   // ---- GENERATED: setup
   IF #Startup OR NOT #Core.Named THEN
       #InstancePath := GetInstancePath(size := 0);
       "FRK_SetIdentity"(Core := #Core,
                         Status := #Status,
                         InstancePath := #InstancePath,
                         ModuleType := 1,
                         TypeId := 4,
                         Capabilities := DWORD#16#00000000,
                         ParentIndex := #ParentIndex,
                         TypeKey := 'Fraktal.Test.Satellite');
   END_IF;
   IF #Startup OR #ConfigRev = 0 THEN
       #ConfigRev := "FRK_ConfigRevision"(Previous := #ConfigRev);
   END_IF;
   #SupportedModesPublished[0] := TRUE;
   #SupportedModesPublished[1] := TRUE;
   #SupportedModesPublished[2] := TRUE;
   #SupportedModesPublished[3] := FALSE;
   #SupportedModesPublished[4] := FALSE;
   #SupportedModesPublished[5] := FALSE;
   #SupportedModesPublished[6] := FALSE;
   "FRK_UnitPrepare"(Core := #Core,
                     Unit := #Unit,
                     Policy := #ModePolicy,
                     Request := #HmiRequest,
                     Response := #HmiResponse,
                     Startup := #Startup,
                     InitialMode := 1);
   "FRK_AccessCyclic"(Access := #Access,
                      Startup := #Startup,
                      SourcePath := STRING_TO_WSTRING(#Status.Name),
                      History := #History,
                      Head := #HistoryHead,
                      Revision := #ConfigRev);
   "FRK_UnitMailbox"(Core := #Core,
                     Unit := #Unit,
                     Status := #Status,
                     Policy := #ModePolicy,
                     Access := #Access,
                     Request := #HmiRequest,
                     Response := #HmiResponse,
                     Supported := #SupportedModesPublished);
   // ---- GENERATED: begin
   "FRK_Begin"(Core := #Core,
               Status := #Status,
               Execute := #Unit.RunReq,
               Abort := (#Abort OR #Unit.AbortReq),
               Command := 1);
   IF #Core.EvCommandStart THEN
       #LatchedParCmd := #ParCmd;
       CASE #Core.Command OF
           1:
               "FRK_UnitRunStart"(Core := #Core,
                                  Status := #Status,
                                  Timeout := #ParCfg.Timeout,
                                  Label := 'Run');
           ELSE
               "FRK_Start"(Core := #Core,
                           Status := #Status,
                           Supported := FALSE,
                           Timeout := T#0ms,
                           Label := '');
       END_CASE;
   END_IF;
   IF #Core.EvCommandStart THEN
       // ---- AUTHORED: CommandStart
       #Device.Received := "FRK_PartReceived"(Core := #Core, Unit := #Unit, Status := #Status, Part := #Part, History := #History, Head := #HistoryHead);
       IF #Device.Received THEN
           "FRK_PartStarted"(Unit := #Unit,
                             Status := #Status,
                             Part := #Part,
                             History := #History,
                             Head := #HistoryHead);
       END_IF;
       // ---- GENERATED: reaction end
   END_IF;
   // ---- AUTHORED: cyclic management
   IF #Hal.Cell.Clamp.BackgroundFault THEN
       "FRK_Fault"(Core := #Core,
                   Status := #Status,
                   ReasonCode := 2901,
                   Description := WSTRING#'test.unit.condition');
   END_IF;
   // ---- GENERATED: end management
   "FRK_Release_SatelliteUnit"(Unit := #Unit,
                               Hal := #Hal);
   "FRK_UnitConsume"(Core := #Core,
                     Unit := #Unit,
                     Status := #Status,
                     Policy := #ModePolicy,
                     Access := #Access,
                     Response := #HmiResponse,
                     Supported := #SupportedModesPublished);
   "FRK_UnitMode"(Core := #Core,
                  Unit := #Unit);
   IF #Core.EvModeExit THEN
       // ---- AUTHORED: ModeExit
       #Device.ExitCalls := #Device.ExitCalls + 1;
       IF #Hal.Cell.Clamp.ExitHold THEN
           #Core.HookResult := 1;
       ELSE
           #Core.HookResult := 0;
       END_IF;
       // ---- GENERATED: reaction end
   END_IF;
   "FRK_UnitModeResolve"(Core := #Core,
                         Unit := #Unit,
                         Status := #Status,
                         Policy := #ModePolicy,
                         Timeout := #ParCfg.Timeout);
   IF #Core.EvModeChanged THEN
       // ---- AUTHORED: ModeChanged
       #Device.Changes := #Device.Changes + 1;
       // ---- GENERATED: reaction end
   END_IF;
   "FRK_UnitFollow"(Core := #Core,
                    Unit := #Unit,
                    Status := #Status,
                    Policy := #ModePolicy,
                    Access := #Access,
                    Supported := #SupportedModesPublished);
   IF #Unit.RequestPending AND (#Unit.Request.Kind = 11 OR #Unit.Request.Kind = 16) THEN
       #ManualMatched := FALSE;
       #RouteMatched := "FRK_Route_DeclarationCell"(Module := #Cell, Hal := #Hal.Cell, Request := #Unit.Request, Report := #HmiResponse.Report);
       #ManualMatched := #ManualMatched OR #RouteMatched;
       #RouteMatched := "FRK_Route_InnerUnit"(Module := #Inner, Hal := #Hal.Inner, Request := #Unit.Request, Report := #HmiResponse.Report);
       #ManualMatched := #ManualMatched OR #RouteMatched;
       IF NOT #ManualMatched THEN
           "FRK_ReleaseReason"(Report := #HmiResponse.Report,
                               Description := WSTRING#'std.error.unsupportedHmiRequest',
                               Reason := 2008,
                               Path := #Unit.Request.TargetPath,
                               Kind := 4);
       END_IF;
       #HmiResponse.Accepted := #Unit.Request.Kind = 16 OR #HmiResponse.Report.Released;
       IF #Unit.Request.Kind = 11 THEN
           IF #HmiResponse.Accepted THEN
               #HmiResponse.Diagnostic := WSTRING#'std.audit.manualCommandAccepted';
           ELSE
               #HmiResponse.Diagnostic := WSTRING#'std.audit.manualCommandRejected';
           END_IF;
       END_IF;
   END_IF;
   IF #Unit.EvReset THEN
       // ---- AUTHORED: OperatorReset
       #Device.Resets := #Device.Resets + 1;
       // ---- GENERATED: reset reaction end
   END_IF;
   IF #Core.ReleasePending OR #Unit.ReleaseChildren THEN
       "FRK_ReleaseCommand"(Core := #Cell.Core,
                            Execute := #Cell.Execute);
       "FRK_ReleaseCommand"(Core := #Inner.Core,
                            Execute := #Inner.Execute);
   END_IF;
   // ---- GENERATED: child call
   #Cell(ParentIndex := #Core.RegIndex,
         Startup := #Startup,
         Hal := #Hal.Cell);
   "FRK_ManualFinish"(Core := #Cell.Core,
                      Execute := #Cell.Execute,
                      ManualOwned := #Cell.ManualOwned);
   "FRK_UnitCascade"(ParentUnit := #Unit,
                     Core := #Inner.Core,
                     Unit := #Inner.Unit,
                     Status := #Inner.Status,
                     Policy := #Inner.ModePolicy,
                     Access := #Inner.Access,
                     Supported := #Inner.SupportedModesPublished,
                     History := #History,
                     Head := #HistoryHead);
   // ---- GENERATED: child call
   #Inner(ParentIndex := #Core.RegIndex,
          Startup := #Startup,
          Hal := #Hal.Inner);
   #Unit.CascadePending := FALSE;
   IF #Unit.RequestPending AND #Unit.Request.Kind = 23 THEN
       #HmiResponse.Accepted := FALSE;
       #HmiResponse.Report.Count := 0;
       #HmiResponse.Report.Released := TRUE;
       #HmiResponse.Diagnostic := WSTRING#'';
       "FRK_ConfigBegin"(Cursor := #ConfigCursor,
                         Page := #HmiResponse.ConfigPage,
                         PageIndex := #Unit.Request.IntValue,
                         Revision := #ConfigRev);
       IF #Unit.Request.DurationMs <> 0 THEN
           #HmiResponse.Diagnostic := WSTRING#'std.error.modelNotAvailable';
       ELSIF #Unit.Request.IntValue < 0 OR #Unit.Request.IntValue > 32767 THEN
           #HmiResponse.Diagnostic := WSTRING#'std.error.hmiRequestRejected';
       ELSE
           "FRK_ConfigUnit"(Scope := #Status.Name,
                            Policy := #ModePolicy,
                            ReadLevel := #Access.Policy.Required[0],
                            Readable := #Access.CurrentLevel >= #Access.Policy.Required[0],
                            Cursor := #ConfigCursor,
                            Page := #HmiResponse.ConfigPage);
           "FRK_Config_DeclarationCell"(Module := #Cell,
                                        ReadLevel := #Access.Policy.Required[0],
                                        Readable := #Access.CurrentLevel >= #Access.Policy.Required[0],
                                        Cursor := #ConfigCursor,
                                        Page := #HmiResponse.ConfigPage);
           "FRK_Config_InnerUnit"(Module := #Inner,
                                  ReadLevel := #Access.Policy.Required[0],
                                  Readable := #Access.CurrentLevel >= #Access.Policy.Required[0],
                                  Cursor := #ConfigCursor,
                                  Page := #HmiResponse.ConfigPage);
           "FRK_ConfigFinish"(Cursor := #ConfigCursor,
                              Page := #HmiResponse.ConfigPage);
           #HmiResponse.Accepted := TRUE;
       END_IF;
   END_IF;
   "FRK_RouteAbort"(Core := #Core,
                    Abort := (#Abort OR #Unit.AbortReq));
   IF #Core.EvAbort THEN
       "FRK_PartAborted"(Core := #Core,
                         Unit := #Unit,
                         Status := #Status,
                         Part := #Part,
                         History := #History,
                         Head := #HistoryHead);
   END_IF;
   IF #Core.Dispatch AND #Core.RegIndex > 0 AND NOT "FRK_Registry".Fault THEN
       // ---- AUTHORED: dispatch
       IF #Hal.Cell.Clamp.Finish THEN
           #Device.Processed := FALSE;
           IF #Unit.CarrierIndex = 0 THEN
               #Device.Processed := TRUE;
           ELSE
               #Device.Processed := "FRK_PartProcessed"(Core := #Core, Unit := #Unit, Status := #Status, Part := #Part, History := #History, Head := #HistoryHead, Verdict := #Hal.Cell.Clamp.Verdict, Reason := #Hal.Cell.Clamp.Diag.ReasonCode);
           END_IF;
           IF #Device.Processed THEN
               #Device.Cycles := #Device.Cycles + 1;
               IF #Unit.StopReq THEN
                   "FRK_Complete"(Core := #Core,
                                  Status := #Status);
               ELSE
                   #Device.Received := "FRK_PartReceived"(Core := #Core, Unit := #Unit, Status := #Status, Part := #Part, History := #History, Head := #HistoryHead);
                   IF #Device.Received THEN
                       "FRK_PartStarted"(Unit := #Unit,
                                         Status := #Status,
                                         Part := #Part,
                                         History := #History,
                                         Head := #HistoryHead);
                   END_IF;
               END_IF;
           END_IF;
       END_IF;
       // ---- GENERATED: end dispatch
   END_IF;
   "FRK_End"(Core := #Core,
             Status := #Status,
             Busy => #Busy,
             Done => #Done,
             Error => #Error,
             Aborted => #Aborted,
             Held => #Held,
             ErrorID => #ErrorID,
             Timing => #Timing);
   "FRK_AccessFinish"(Access := #Access,
                      Unit := #Unit,
                      Response := #HmiResponse,
                      SourcePath := STRING_TO_WSTRING(#Status.Name),
                      History := #History,
                      Head := #HistoryHead,
                      Revision := #ConfigRev);
   "FRK_UnitFinish"(Core := #Core,
                    Unit := #Unit,
                    Response := #HmiResponse,
                    Status := #Status,
                    Part := #Part,
                    History := #History,
                    Head := #HistoryHead);
   #ModeActivePublished := #Unit.Mode;
   #RunningPublished := #Core.Exec = 1;
   #StopPendingPublished := #Unit.StopReq AND #Core.Exec = 1;
   #GoodCount := #Unit.Good;
   #NokCount := #Unit.Nok;
   #ReworkCount := #Unit.Rework;
   #NokReason := #Unit.NokReason;
   // ---- AUTHORED: unconditional cyclic/derived data
   #OutImm.Cycles := #Device.Cycles;
   #OutImm.ExitCalls := #Device.ExitCalls;
   #OutImm.Changes := #Device.Changes;
   #OutImm.Resets := #Device.Resets;
   // ---- GENERATED: frame end
END_FUNCTION_BLOCK

FUNCTION_BLOCK "FB_InnerUnit"   // FB3, SCL
{ S7_Optimized_Access := 'TRUE' }
VERSION : 0.1
// Generated frame v0.6; change the declaration, then regenerate.
// stored: AutoNumber true, IsIECCheckEnabled false, IsRetainMemResEnabled false, MemoryReserve 100, SetENOAutomatically false, UDAEnableTagReadback false
   VAR_INPUT
      Execute { ExternalWritable := 'False'} : Bool;
      Abort { ExternalWritable := 'False'} : Bool;
      Command { ExternalWritable := 'False'} : DInt;
      ParCfg { ExternalWritable := 'False'} : "ST_DeclarationParCfg";
      ParCmd { ExternalWritable := 'False'} : "ST_DeclarationParCmd";
      ParentIndex { ExternalAccessible := 'False'; ExternalVisible := 'False'; ExternalWritable := 'False'} : DInt;
      Startup { ExternalAccessible := 'False'; ExternalVisible := 'False'; ExternalWritable := 'False'} : Bool;
   END_VAR
   VAR_OUTPUT
      Busy { ExternalWritable := 'False'} : Bool;
      Done { ExternalWritable := 'False'} : Bool;
      Error { ExternalWritable := 'False'} : Bool;
      Aborted { ExternalWritable := 'False'} : Bool;
      Held { ExternalWritable := 'False'} : Bool;
      ErrorID { ExternalWritable := 'False'} : DWord;
      Timing { ExternalWritable := 'False'} : "ST_ModuleTiming";
      OutCmd { ExternalWritable := 'False'} : "ST_DeclarationOutCmd";
      OutImm { ExternalWritable := 'False'} : "ST_UnitProbeImm";
   END_VAR
   VAR_IN_OUT
      Hal : "ST_InnerUnitHal";
   END_VAR
   VAR
      Status { ExternalWritable := 'False'; S7_SetPoint := 'True'} : "ST_ModuleStatus";
      Core { ExternalAccessible := 'False'; ExternalVisible := 'False'; ExternalWritable := 'False'; S7_SetPoint := 'True'} : "FRK_Core";
      LatchedParCmd { ExternalAccessible := 'False'; ExternalVisible := 'False'; ExternalWritable := 'False'; S7_SetPoint := 'True'} : "ST_DeclarationParCmd";
      Device { ExternalAccessible := 'False'; ExternalVisible := 'False'; ExternalWritable := 'False'; S7_SetPoint := 'True'} : "ST_UnitProbeDevice";
      Unit { ExternalAccessible := 'False'; ExternalVisible := 'False'; ExternalWritable := 'False'; S7_SetPoint := 'True'} : "FRK_Unit";
      HmiRequest { S7_SetPoint := 'True'} : "ST_HmiRequest";
      ModePolicy { ExternalAccessible := 'False'; ExternalVisible := 'False'; ExternalWritable := 'False'; S7_SetPoint := 'True'} : Array[0..6] of "ST_ModePolicy";
      Access { ExternalWritable := 'False'; S7_SetPoint := 'True'} : "FRK_Access";
      HmiResponse { ExternalWritable := 'False'; S7_SetPoint := 'True'} : "ST_HmiResponse";
      ConfigRev { ExternalWritable := 'False'} : UDInt;
      ConfigCursor { ExternalAccessible := 'False'; ExternalVisible := 'False'; ExternalWritable := 'False'; S7_SetPoint := 'True'} : "FRK_ConfigCursor";
      Part { ExternalWritable := 'False'; S7_SetPoint := 'True'} : "ST_PartContext";
      History { ExternalWritable := 'False'; S7_SetPoint := 'True'} : Array[1..16] of "ST_Diagnostic";
      HistoryHead { ExternalWritable := 'False'} : Int;
      ModeActivePublished { ExternalWritable := 'False'} : DInt;
      RunningPublished { ExternalWritable := 'False'} : Bool;
      StopPendingPublished { ExternalWritable := 'False'} : Bool;
      SupportedModesPublished { ExternalWritable := 'False'} : Array[0..6] of Bool;
      GoodCount { ExternalWritable := 'False'} : UDInt;
      NokCount { ExternalWritable := 'False'} : UDInt;
      ReworkCount { ExternalWritable := 'False'} : UDInt;
      NokReason { ExternalWritable := 'False'} : DInt;
      Cell { ExternalWritable := 'False'; S7_SetPoint := 'True'} : "FB_DeclarationCell";
   END_VAR
   VAR_TEMP
      InstancePath : WString[254];
      RouteMatched : Bool;
      ManualMatched : Bool;
   END_VAR
   VAR CONSTANT
      EXEC_READY : DInt := 0;
      MODULE_TIER : DInt := 1;
   END_VAR
BEGIN

   // ---- GENERATED: setup
   IF #Startup OR NOT #Core.Named THEN
       #InstancePath := GetInstancePath(size := 0);
       "FRK_SetIdentity"(Core := #Core,
                         Status := #Status,
                         InstancePath := #InstancePath,
                         ModuleType := 1,
                         TypeId := 5,
                         Capabilities := DWORD#16#00000000,
                         ParentIndex := #ParentIndex,
                         TypeKey := 'Fraktal.Test.Inner');
   END_IF;
   IF #Startup OR #ConfigRev = 0 THEN
       #ConfigRev := "FRK_ConfigRevision"(Previous := #ConfigRev);
   END_IF;
   #SupportedModesPublished[0] := TRUE;
   #SupportedModesPublished[1] := TRUE;
   #SupportedModesPublished[2] := TRUE;
   #SupportedModesPublished[3] := FALSE;
   #SupportedModesPublished[4] := FALSE;
   #SupportedModesPublished[5] := FALSE;
   #SupportedModesPublished[6] := FALSE;
   "FRK_UnitPrepare"(Core := #Core,
                     Unit := #Unit,
                     Policy := #ModePolicy,
                     Request := #HmiRequest,
                     Response := #HmiResponse,
                     Startup := #Startup,
                     InitialMode := 1);
   "FRK_AccessCyclic"(Access := #Access,
                      Startup := #Startup,
                      SourcePath := STRING_TO_WSTRING(#Status.Name),
                      History := #History,
                      Head := #HistoryHead,
                      Revision := #ConfigRev);
   "FRK_UnitMailbox"(Core := #Core,
                     Unit := #Unit,
                     Status := #Status,
                     Policy := #ModePolicy,
                     Access := #Access,
                     Request := #HmiRequest,
                     Response := #HmiResponse,
                     Supported := #SupportedModesPublished);
   // ---- GENERATED: begin
   "FRK_Begin"(Core := #Core,
               Status := #Status,
               Execute := #Unit.RunReq,
               Abort := (#Abort OR #Unit.AbortReq),
               Command := 1);
   IF #Core.EvCommandStart THEN
       #LatchedParCmd := #ParCmd;
       CASE #Core.Command OF
           1:
               "FRK_UnitRunStart"(Core := #Core,
                                  Status := #Status,
                                  Timeout := #ParCfg.Timeout,
                                  Label := 'Run');
           ELSE
               "FRK_Start"(Core := #Core,
                           Status := #Status,
                           Supported := FALSE,
                           Timeout := T#0ms,
                           Label := '');
       END_CASE;
   END_IF;
   IF #Core.EvCommandStart THEN
       // ---- AUTHORED: CommandStart
       #Device.Received := "FRK_PartReceived"(Core := #Core, Unit := #Unit, Status := #Status, Part := #Part, History := #History, Head := #HistoryHead);
       IF #Device.Received THEN
           "FRK_PartStarted"(Unit := #Unit,
                             Status := #Status,
                             Part := #Part,
                             History := #History,
                             Head := #HistoryHead);
       END_IF;
       // ---- GENERATED: reaction end
   END_IF;
   // ---- AUTHORED: cyclic management
   IF #Hal.Cell.Clamp.BackgroundFault THEN
       "FRK_Fault"(Core := #Core,
                   Status := #Status,
                   ReasonCode := 2901,
                   Description := WSTRING#'test.unit.condition');
   END_IF;
   // ---- GENERATED: end management
   "FRK_Release_InnerUnit"(Unit := #Unit,
                           Hal := #Hal);
   "FRK_UnitConsume"(Core := #Core,
                     Unit := #Unit,
                     Status := #Status,
                     Policy := #ModePolicy,
                     Access := #Access,
                     Response := #HmiResponse,
                     Supported := #SupportedModesPublished);
   "FRK_UnitMode"(Core := #Core,
                  Unit := #Unit);
   IF #Core.EvModeExit THEN
       // ---- AUTHORED: ModeExit
       #Device.ExitCalls := #Device.ExitCalls + 1;
       IF #Hal.Cell.Clamp.ExitHold THEN
           #Core.HookResult := 1;
       ELSE
           #Core.HookResult := 0;
       END_IF;
       // ---- GENERATED: reaction end
   END_IF;
   "FRK_UnitModeResolve"(Core := #Core,
                         Unit := #Unit,
                         Status := #Status,
                         Policy := #ModePolicy,
                         Timeout := #ParCfg.Timeout);
   IF #Core.EvModeChanged THEN
       // ---- AUTHORED: ModeChanged
       #Device.Changes := #Device.Changes + 1;
       // ---- GENERATED: reaction end
   END_IF;
   "FRK_UnitFollow"(Core := #Core,
                    Unit := #Unit,
                    Status := #Status,
                    Policy := #ModePolicy,
                    Access := #Access,
                    Supported := #SupportedModesPublished);
   IF #Unit.RequestPending AND (#Unit.Request.Kind = 11 OR #Unit.Request.Kind = 16) THEN
       #ManualMatched := FALSE;
       #RouteMatched := "FRK_Route_DeclarationCell"(Module := #Cell, Hal := #Hal.Cell, Request := #Unit.Request, Report := #HmiResponse.Report);
       #ManualMatched := #ManualMatched OR #RouteMatched;
       IF NOT #ManualMatched THEN
           "FRK_ReleaseReason"(Report := #HmiResponse.Report,
                               Description := WSTRING#'std.error.unsupportedHmiRequest',
                               Reason := 2008,
                               Path := #Unit.Request.TargetPath,
                               Kind := 4);
       END_IF;
       #HmiResponse.Accepted := #Unit.Request.Kind = 16 OR #HmiResponse.Report.Released;
       IF #Unit.Request.Kind = 11 THEN
           IF #HmiResponse.Accepted THEN
               #HmiResponse.Diagnostic := WSTRING#'std.audit.manualCommandAccepted';
           ELSE
               #HmiResponse.Diagnostic := WSTRING#'std.audit.manualCommandRejected';
           END_IF;
       END_IF;
   END_IF;
   IF #Unit.EvReset THEN
       // ---- AUTHORED: OperatorReset
       #Device.Resets := #Device.Resets + 1;
       // ---- GENERATED: reset reaction end
   END_IF;
   IF #Core.ReleasePending OR #Unit.ReleaseChildren THEN
       "FRK_ReleaseCommand"(Core := #Cell.Core,
                            Execute := #Cell.Execute);
   END_IF;
   // ---- GENERATED: child call
   #Cell(ParentIndex := #Core.RegIndex,
         Startup := #Startup,
         Hal := #Hal.Cell);
   "FRK_ManualFinish"(Core := #Cell.Core,
                      Execute := #Cell.Execute,
                      ManualOwned := #Cell.ManualOwned);
   #Unit.CascadePending := FALSE;
   IF #Unit.RequestPending AND #Unit.Request.Kind = 23 THEN
       #HmiResponse.Accepted := FALSE;
       #HmiResponse.Report.Count := 0;
       #HmiResponse.Report.Released := TRUE;
       #HmiResponse.Diagnostic := WSTRING#'';
       "FRK_ConfigBegin"(Cursor := #ConfigCursor,
                         Page := #HmiResponse.ConfigPage,
                         PageIndex := #Unit.Request.IntValue,
                         Revision := #ConfigRev);
       IF #Unit.Request.DurationMs <> 0 THEN
           #HmiResponse.Diagnostic := WSTRING#'std.error.modelNotAvailable';
       ELSIF #Unit.Request.IntValue < 0 OR #Unit.Request.IntValue > 32767 THEN
           #HmiResponse.Diagnostic := WSTRING#'std.error.hmiRequestRejected';
       ELSE
           "FRK_ConfigUnit"(Scope := #Status.Name,
                            Policy := #ModePolicy,
                            ReadLevel := #Access.Policy.Required[0],
                            Readable := #Access.CurrentLevel >= #Access.Policy.Required[0],
                            Cursor := #ConfigCursor,
                            Page := #HmiResponse.ConfigPage);
           "FRK_Config_DeclarationCell"(Module := #Cell,
                                        ReadLevel := #Access.Policy.Required[0],
                                        Readable := #Access.CurrentLevel >= #Access.Policy.Required[0],
                                        Cursor := #ConfigCursor,
                                        Page := #HmiResponse.ConfigPage);
           "FRK_ConfigFinish"(Cursor := #ConfigCursor,
                              Page := #HmiResponse.ConfigPage);
           #HmiResponse.Accepted := TRUE;
       END_IF;
   END_IF;
   "FRK_RouteAbort"(Core := #Core,
                    Abort := (#Abort OR #Unit.AbortReq));
   IF #Core.EvAbort THEN
       "FRK_PartAborted"(Core := #Core,
                         Unit := #Unit,
                         Status := #Status,
                         Part := #Part,
                         History := #History,
                         Head := #HistoryHead);
   END_IF;
   IF #Core.Dispatch AND #Core.RegIndex > 0 AND NOT "FRK_Registry".Fault THEN
       // ---- AUTHORED: dispatch
       IF #Hal.Cell.Clamp.Finish THEN
           #Device.Processed := FALSE;
           IF #Unit.CarrierIndex = 0 THEN
               #Device.Processed := TRUE;
           ELSE
               #Device.Processed := "FRK_PartProcessed"(Core := #Core, Unit := #Unit, Status := #Status, Part := #Part, History := #History, Head := #HistoryHead, Verdict := #Hal.Cell.Clamp.Verdict, Reason := #Hal.Cell.Clamp.Diag.ReasonCode);
           END_IF;
           IF #Device.Processed THEN
               #Device.Cycles := #Device.Cycles + 1;
               IF #Unit.StopReq THEN
                   "FRK_Complete"(Core := #Core,
                                  Status := #Status);
               ELSE
                   #Device.Received := "FRK_PartReceived"(Core := #Core, Unit := #Unit, Status := #Status, Part := #Part, History := #History, Head := #HistoryHead);
                   IF #Device.Received THEN
                       "FRK_PartStarted"(Unit := #Unit,
                                         Status := #Status,
                                         Part := #Part,
                                         History := #History,
                                         Head := #HistoryHead);
                   END_IF;
               END_IF;
           END_IF;
       END_IF;
       // ---- GENERATED: end dispatch
   END_IF;
   "FRK_End"(Core := #Core,
             Status := #Status,
             Busy => #Busy,
             Done => #Done,
             Error => #Error,
             Aborted => #Aborted,
             Held => #Held,
             ErrorID => #ErrorID,
             Timing => #Timing);
   "FRK_AccessFinish"(Access := #Access,
                      Unit := #Unit,
                      Response := #HmiResponse,
                      SourcePath := STRING_TO_WSTRING(#Status.Name),
                      History := #History,
                      Head := #HistoryHead,
                      Revision := #ConfigRev);
   "FRK_UnitFinish"(Core := #Core,
                    Unit := #Unit,
                    Response := #HmiResponse,
                    Status := #Status,
                    Part := #Part,
                    History := #History,
                    Head := #HistoryHead);
   #ModeActivePublished := #Unit.Mode;
   #RunningPublished := #Core.Exec = 1;
   #StopPendingPublished := #Unit.StopReq AND #Core.Exec = 1;
   #GoodCount := #Unit.Good;
   #NokCount := #Unit.Nok;
   #ReworkCount := #Unit.Rework;
   #NokReason := #Unit.NokReason;
   // ---- AUTHORED: unconditional cyclic/derived data
   #OutImm.Cycles := #Device.Cycles;
   #OutImm.ExitCalls := #Device.ExitCalls;
   #OutImm.Changes := #Device.Changes;
   #OutImm.Resets := #Device.Resets;
   // ---- GENERATED: frame end
END_FUNCTION_BLOCK

FUNCTION "FRK_AccessAudit" : Void   // FC32, SCL
{ S7_Optimized_Access := 'TRUE' }
VERSION : 0.1
// stored: AutoNumber true, IsIECCheckEnabled false, SetENOAutomatically false, UDAEnableTagReadback false
   VAR_INPUT
      What : WString;
      Who : String;
      SourcePath : WString;
   END_VAR
   VAR_IN_OUT
      History : Array[1..16] of "ST_Diagnostic";
      Head : Int;
   END_VAR
   VAR_TEMP
      Description : WString[480];
   END_VAR
BEGIN

   #Description := CONCAT(IN1 := #What, IN2 := WSTRING#': ');
   #Description := CONCAT(IN1 := #Description, IN2 := STRING_TO_WSTRING(#Who));
   "FRK_HistoryEvent"(History := #History,
                      Head := #Head,
                      Reason := 0,
                      Description := #Description,
                      SourcePath := #SourcePath);
END_FUNCTION

FUNCTION "FRK_AccessCancel" : Void   // FC27, SCL
{ S7_Optimized_Access := 'TRUE' }
VERSION : 0.1
// stored: AutoNumber true, IsIECCheckEnabled false, SetENOAutomatically false, UDAEnableTagReadback false
   VAR_IN_OUT
      Access : "FRK_Access";
   END_VAR
   VAR_TEMP
      Index : DInt;
   END_VAR
BEGIN

   #Access.LoginBusy := FALSE;
   #Access.CandidateUser := '';
   #Access.CandidateLevel := 0;
   #Access.Round := 0;
   FOR #Index := 0 TO 15 DO
       #Access.Salt[#Index] := 0;
   END_FOR;
   FOR #Index := 0 TO 31 DO
       #Access.Digest[#Index] := 0;
       #Access.Expected[#Index] := 0;
   END_FOR;
END_FUNCTION

FUNCTION "FRK_AccessCyclic" : Void   // FC33, SCL
{ S7_Optimized_Access := 'TRUE' }
VERSION : 0.1
// stored: AutoNumber true, IsIECCheckEnabled false, SetENOAutomatically false, UDAEnableTagReadback false
   VAR_INPUT
      Startup : Bool;
      SourcePath : WString;
   END_VAR
   VAR_IN_OUT
      Access : "FRK_Access";
      History : Array[1..16] of "ST_Diagnostic";
      Head : Int;
      Revision : UDInt;
   END_VAR
   VAR_TEMP
      Data : Array[0..47] of Byte;
      Index : DInt;
      Difference : Byte;
      HashOk : Bool;
   END_VAR
BEGIN

   #Access.LoginTimeoutMs := 6000;
   IF #Startup THEN
       "FRK_AccessLogout"(Access := #Access);
       #Access.LoginResultSequence := 0;
   END_IF;
   IF #Access.CurrentLevel > 0 AND #Access.Policy.SessionTimeout > T#0ms THEN
       IF "FRK_Elapsed"(NewMs := "FRK_Clock".NowMs, OldMs := #Access.LastActivity) >= DINT_TO_UDINT(TIME_TO_DINT(#Access.Policy.SessionTimeout)) THEN
           "FRK_AccessAudit"(History := #History,
                             Head := #Head,
                             What := WSTRING#'std.audit.autoLogout',
                             Who := #Access.CurrentUser,
                             SourcePath := #SourcePath);
           // Expiring the old session does not discard a separately committed
           // credential attempt. Explicit logout cancels both.
           "FRK_AccessDropSession"(Access := #Access);
           #Revision := "FRK_ConfigRevision"(Previous := #Revision);
       END_IF;
   END_IF;
   IF NOT #Access.LoginBusy THEN
       RETURN;
   END_IF;
   // One compression per active scan; never run all PIN rounds in one scan.
   FOR #Index := 0 TO 31 DO
       #Data[#Index] := #Access.Digest[#Index];
   END_FOR;
   FOR #Index := 0 TO 15 DO
       #Data[32 + #Index] := #Access.Salt[#Index];
   END_FOR;
   #HashOk := "FRK_Sha256Pin"(Data := #Data, Size := 48, Digest := #Access.Digest);
   FOR #Index := 0 TO 47 DO
       #Data[#Index] := 0;
   END_FOR;
   #Access.Round := #Access.Round + 1;
   IF NOT #HashOk OR "FRK_Elapsed"(NewMs := "FRK_Clock".NowMs, OldMs := #Access.LoginSince) >= #Access.LoginTimeoutMs THEN
       #Access.CandidateLevel := 0;
   ELSIF #Access.Round < 256 THEN
       RETURN;
   END_IF;
   #Difference := 0;
   FOR #Index := 0 TO 31 DO
       #Difference := #Difference OR (#Access.Digest[#Index] XOR #Access.Expected[#Index]);
   END_FOR;
   #Access.LoginFailed := #Difference <> 0 OR #Access.CandidateLevel = 0 OR NOT #Access.ProviderEnabled;
   IF #Access.LoginFailed THEN
       "FRK_AccessAudit"(History := #History,
                         Head := #Head,
                         What := WSTRING#'std.audit.loginFailed',
                         Who := #Access.CandidateUser,
                         SourcePath := #SourcePath);
   ELSE
       #Access.CurrentUser := #Access.CandidateUser;
       #Access.CurrentLevel := #Access.CandidateLevel;
       #Access.LastActivity := "FRK_Clock".NowMs;
       #Access.SessionGeneration := "FRK_AccessNext"(Previous := #Access.SessionGeneration);
       #Revision := "FRK_ConfigRevision"(Previous := #Revision);
       "FRK_AccessAudit"(History := #History,
                         Head := #Head,
                         What := WSTRING#'std.audit.login',
                         Who := #Access.CurrentUser,
                         SourcePath := #SourcePath);
   END_IF;
   #Access.LoginResultSequence := #Access.LoginSequence;
   "FRK_AccessCancel"(Access := #Access);
END_FUNCTION

FUNCTION "FRK_AccessDropSession" : Void   // FC29, SCL
{ S7_Optimized_Access := 'TRUE' }
VERSION : 0.1
// stored: AutoNumber true, IsIECCheckEnabled false, SetENOAutomatically false, UDAEnableTagReadback false
   VAR_IN_OUT
      Access : "FRK_Access";
   END_VAR
BEGIN

   #Access.CurrentLevel := 0;
   #Access.CurrentUser := '';
   #Access.LoginFailed := FALSE;
   #Access.SessionGeneration := "FRK_AccessNext"(Previous := #Access.SessionGeneration);
END_FUNCTION

FUNCTION "FRK_AccessFinish" : Void   // FC34, SCL
{ S7_Optimized_Access := 'TRUE' }
VERSION : 0.1
// stored: AutoNumber true, IsIECCheckEnabled false, SetENOAutomatically false, UDAEnableTagReadback false
   VAR_INPUT
      Unit : "FRK_Unit";
      Response : "ST_HmiResponse";
      SourcePath : WString;
   END_VAR
   VAR_IN_OUT
      Access : "FRK_Access";
      History : Array[1..16] of "ST_Diagnostic";
      Head : Int;
      Revision : UDInt;
   END_VAR
   VAR_TEMP
      What : WString[160];
      AuditPath : WString[255];
   END_VAR
BEGIN

   IF NOT #Unit.RequestPending THEN
       RETURN;
   END_IF;
   CASE #Unit.Request.Kind OF
       23, 15,
       16, 17,
       1:
           RETURN;
       2:
           "FRK_AccessAudit"(History := #History,
                             Head := #Head,
                             What := WSTRING#'std.audit.logout',
                             Who := #Unit.RequestUser,
                             SourcePath := #SourcePath);
           #Revision := "FRK_ConfigRevision"(Previous := #Revision);
           RETURN;
       ELSE
           #What := WSTRING#'std.audit.accessDenied';
   END_CASE;
   IF #Response.Accepted THEN
       #What := WSTRING#'std.audit.operatorAction';
       IF #Access.CurrentLevel > 0 THEN
           #Access.LastActivity := "FRK_Clock".NowMs;
       END_IF;
       IF #Unit.Request.Kind = 24 THEN
           #Revision := "FRK_ConfigRevision"(Previous := #Revision);
       END_IF;
   END_IF;
   #AuditPath := #SourcePath;
   IF #Unit.Request.Kind = 11 THEN
       #AuditPath := #Unit.Request.TargetPath;
       IF #Response.Accepted THEN
           #What := WSTRING#'std.audit.manualCommandAccepted';
       ELSE
           #What := WSTRING#'std.audit.manualCommandRejected';
       END_IF;
   END_IF;
   #What := CONCAT(IN1 := #What, IN2 := WSTRING#' kind=');
   #What := CONCAT(IN1 := #What, IN2 := DINT_TO_WSTRING(#Unit.Request.Kind));
   #What := CONCAT(IN1 := #What, IN2 := WSTRING#' value=');
   #What := CONCAT(IN1 := #What, IN2 := DINT_TO_WSTRING(#Unit.Request.IntValue));
   "FRK_AccessAudit"(History := #History,
                     Head := #Head,
                     What := #What,
                     Who := #Unit.RequestUser,
                     SourcePath := #AuditPath);
END_FUNCTION

FUNCTION "FRK_AccessLogin" : Void   // FC31, SCL
{ S7_Optimized_Access := 'TRUE' }
VERSION : 0.1
// stored: AutoNumber true, IsIECCheckEnabled false, SetENOAutomatically false, UDAEnableTagReadback false
   VAR_INPUT
      User : String;
      Secret : String;
      Sequence : UDInt;
   END_VAR
   VAR_IN_OUT
      Access : "FRK_Access";
   END_VAR
   VAR_TEMP
      Data : Array[0..47] of Byte;
      Index : DInt;
      Slot : DInt;
      Size : Int;
      HashOk : Bool;
   END_VAR
BEGIN

   "FRK_AccessCancel"(Access := #Access);
   #Access.LoginFailed := FALSE;
   #Access.LoginSequence := #Sequence;
   #Access.LoginSince := "FRK_Clock".NowMs;
   #Access.LoginTimeoutMs := 6000;
   #Access.CandidateUser := #User;
   // Unknown users execute the same bounded work with a dummy salt/digest.
   IF #Access.ProviderEnabled AND "FRK_LocalUsers".Count >= 0 AND "FRK_LocalUsers".Count <= 16 THEN
       FOR #Slot := 1 TO "FRK_LocalUsers".Count DO
           IF #User <> '' AND "FRK_LocalUsers".Rows[#Slot].User = #User THEN
               IF "FRK_LocalUsers".Rows[#Slot].Level >= 1 AND "FRK_LocalUsers".Rows[#Slot].Level <= 4 THEN
                   #Access.CandidateLevel := "FRK_LocalUsers".Rows[#Slot].Level;
                   #Access.Salt := "FRK_LocalUsers".Rows[#Slot].Salt;
                   #Access.Expected := "FRK_LocalUsers".Rows[#Slot].PinHash;
               END_IF;
               EXIT;
           END_IF;
       END_FOR;
   END_IF;
   FOR #Index := 0 TO 47 DO
       #Data[#Index] := 0;
   END_FOR;
   FOR #Index := 0 TO 15 DO
       #Data[#Index] := #Access.Salt[#Index];
   END_FOR;
   #Size := LEN(#Secret);
   IF #Size > 32 THEN
       #Size := 0;
       #Access.CandidateLevel := 0;
   END_IF;
   FOR #Index := 1 TO #Size DO
       #Data[15 + #Index] := CHAR_TO_BYTE(#Secret[#Index]);
   END_FOR;
   #HashOk := "FRK_Sha256Pin"(Data := #Data, Size := 16 + INT_TO_DINT(#Size), Digest := #Access.Digest);
   FOR #Index := 0 TO 47 DO
       #Data[#Index] := 0;
   END_FOR;
   #Access.LoginBusy := #HashOk;
END_FUNCTION

FUNCTION "FRK_AccessLogout" : Void   // FC28, SCL
{ S7_Optimized_Access := 'TRUE' }
VERSION : 0.1
// stored: AutoNumber true, IsIECCheckEnabled false, SetENOAutomatically false, UDAEnableTagReadback false
   VAR_IN_OUT
      Access : "FRK_Access";
   END_VAR
BEGIN

   "FRK_AccessCancel"(Access := #Access);
   "FRK_AccessDropSession"(Access := #Access);
END_FUNCTION

FUNCTION "FRK_AccessNext" : UDInt   // FC30, SCL
{ S7_Optimized_Access := 'TRUE' }
VERSION : 0.1
// stored: AutoNumber true, IsIECCheckEnabled false, SetENOAutomatically false, UDAEnableTagReadback false
   VAR_INPUT
      Previous : UDInt;
   END_VAR
BEGIN

   IF #Previous = UDINT#4294967295 THEN
       #FRK_AccessNext := 1;
   ELSE
       #FRK_AccessNext := #Previous + 1;
   END_IF;
END_FUNCTION

FUNCTION "FRK_AdoptFault" : Void   // FC9, SCL
{ S7_Optimized_Access := 'TRUE' }
VERSION : 0.1
// stored: AutoNumber true, IsIECCheckEnabled false, SetENOAutomatically false, UDAEnableTagReadback false
   VAR_INPUT
      Diag : "ST_Diagnostic";
   END_VAR
   VAR_IN_OUT
      Core : "FRK_Core";
      Status : "ST_ModuleStatus";
   END_VAR
BEGIN

   IF #Core.Exec = 3 THEN
       RETURN;
   END_IF;
   #Status.Diagnostic := #Diag;
   #Core.Exec := 3;
   #Core.Step := 0;
   #Core.Dispatch := FALSE;
   #Core.DiagTouched := TRUE;
END_FUNCTION

FUNCTION "FRK_Begin" : Void   // FC15, SCL
{ S7_Optimized_Access := 'TRUE' }
VERSION : 0.1
// stored: AutoNumber true, IsIECCheckEnabled false, SetENOAutomatically false, UDAEnableTagReadback false
   VAR_INPUT
      Execute : Bool;
      Abort : Bool;
      Command : DInt;
   END_VAR
   VAR_IN_OUT
      Core : "FRK_Core";
      Status : "ST_ModuleStatus";
   END_VAR
BEGIN

   #Core.EvInit := NOT #Core.Initialized;
   #Core.Initialized := TRUE;
   #Core.EvCommandStart := FALSE;
   #Core.EvAbort := FALSE;
   #Core.EvAbortInError := FALSE;
   #Core.HoldReq := FALSE;
   #Core.DiagTouched := FALSE;
   #Core.HookResult := 0;
   IF NOT #Execute AND (#Core.Armed OR #Core.ReleasePending) AND (#Core.Exec = 2 OR #Core.Exec = 3 OR #Core.Exec = 4) THEN
       #Core.Exec := 0;
       #Core.Armed := FALSE;
       #Core.HoldReason := 0;
       "FRK_ClearDiag"(Status := #Status);
   END_IF;
   IF #Execute AND NOT #Core.ExecPrev AND (#Core.Exec = 0 OR (#Core.Exec = 3 AND NOT #Core.Armed)) THEN
       #Core.Exec := 1;
       #Core.Armed := TRUE;
       #Core.Command := #Command;
       #Core.Step := 10;
       #Core.StartMs := "FRK_Clock".NowMs;
       #Core.LastNowMs := "FRK_Clock".NowMs;
       #Core.ActiveMs := 0;
       #Core.TimeoutMs := 0;
       #Core.CommandLabel := '';
       #Core.TimingOpen := TRUE;
       #Core.Held := FALSE;
       #Core.HoldReason := 0;
       "FRK_ClearDiag"(Status := #Status);
       #Core.EvCommandStart := TRUE;
   END_IF;
   #Core.DeltaMs := "FRK_Elapsed"(NewMs := "FRK_Clock".NowMs, OldMs := #Core.LastNowMs);
   #Core.LastNowMs := "FRK_Clock".NowMs;
   #Core.ExecPrev := #Execute;
   #Core.Dispatch := #Core.Exec = 1;
END_FUNCTION

FUNCTION "FRK_ClearDiag" : Void   // FC5, SCL
{ S7_Optimized_Access := 'TRUE' }
VERSION : 0.1
// stored: AutoNumber true, IsIECCheckEnabled false, SetENOAutomatically false, UDAEnableTagReadback false
   VAR_IN_OUT
      Status : "ST_ModuleStatus";
   END_VAR
BEGIN

   #Status.Diagnostic.ReasonCode := 0;
   #Status.Diagnostic.SourcePath := WSTRING#'';
   #Status.Diagnostic.Description := WSTRING#'';
   #Status.Diagnostic.IoTag := '';
   #Status.Diagnostic.IoAddress := '';
   #Status.Diagnostic.Severity := 0;
   #Status.Diagnostic.Category := 0;
   #Status.Diagnostic.Since := LDT#1970-01-01-00:00:00.000000000;
   #Status.Diagnostic.TimeSynchronized := FALSE;
END_FUNCTION

FUNCTION "FRK_ClockTick" : Void   // FC3, SCL
{ S7_Optimized_Access := 'TRUE' }
VERSION : 0.1
// Shared command kernel v0.1. Core 2.2 / 6.1 / 3.14 / 8.11.
//  Generated enum/rationalization values come from Core authorities.
// stored: AutoNumber true, IsIECCheckEnabled false, SetENOAutomatically false, UDAEnableTagReadback false
   VAR_TEMP
      DeltaS : LReal;
   END_VAR
BEGIN

   #DeltaS := RUNTIME("FRK_Clock".Mem);
   IF #DeltaS < 0.0 OR #DeltaS > 60.0 THEN
       #DeltaS := 0.0;
   END_IF;
   "FRK_Clock".AccMs := "FRK_Clock".AccMs + #DeltaS * 1000.0;
   IF "FRK_Clock".AccMs >= 4294967296.0 THEN
       "FRK_Clock".AccMs := "FRK_Clock".AccMs - 4294967296.0;
   END_IF;
   "FRK_Clock".NowMs := TRUNC_UDINT("FRK_Clock".AccMs);
END_FUNCTION

FUNCTION "FRK_Complete" : Void   // FC13, SCL
{ S7_Optimized_Access := 'TRUE' }
VERSION : 0.1
// stored: AutoNumber true, IsIECCheckEnabled false, SetENOAutomatically false, UDAEnableTagReadback false
   VAR_IN_OUT
      Core : "FRK_Core";
      Status : "ST_ModuleStatus";
   END_VAR
BEGIN

   IF #Core.Exec = 1 THEN
       #Core.Exec := 2;
       #Core.Step := 0;
       #Core.Dispatch := FALSE;
       "FRK_ClearDiag"(Status := #Status);
   END_IF;
END_FUNCTION

FUNCTION "FRK_ConfigAppend" : Void   // FC22, SCL
{ S7_Optimized_Access := 'TRUE' }
VERSION : 0.1
// stored: AutoNumber true, IsIECCheckEnabled false, SetENOAutomatically false, UDAEnableTagReadback false
   VAR_INPUT
      Scope : String;
      Item : String;
      ValueText : WString;
      ValueType : DInt;
      ReadLevel : DInt;
      Readable : Bool;
   END_VAR
   VAR_IN_OUT
      Cursor : "FRK_ConfigCursor";
      Page : "ST_ConfigPage";
   END_VAR
   VAR_TEMP
      Slot : DInt;
   END_VAR
BEGIN

   #Slot := #Cursor.Position - #Cursor.First;
   #Cursor.Position := #Cursor.Position + 1;
   IF #Slot < 0 OR #Slot >= 16 THEN
       RETURN;
   END_IF;
   #Slot := #Slot + 1;
   #Page.Entries[#Slot].Scope := STRING_TO_WSTRING(#Scope);
   #Page.Entries[#Slot].Item := STRING_TO_WSTRING(#Item);
   #Page.Entries[#Slot].ValueType := #ValueType;
   #Page.Entries[#Slot].ReadLevel := #ReadLevel;
   #Page.Entries[#Slot].Readable := #Readable;
   IF #Readable THEN
       #Page.Entries[#Slot].ValueText := #ValueText;
   END_IF;
   #Page.EntryCount := DINT_TO_INT(#Slot);
END_FUNCTION

FUNCTION "FRK_ConfigBegin" : Void   // FC21, SCL
{ S7_Optimized_Access := 'TRUE' }
VERSION : 0.1
// stored: AutoNumber true, IsIECCheckEnabled false, SetENOAutomatically false, UDAEnableTagReadback false
   VAR_INPUT
      PageIndex : DInt;
      Revision : UDInt;
   END_VAR
   VAR_IN_OUT
      Cursor : "FRK_ConfigCursor";
      Page : "ST_ConfigPage";
   END_VAR
   VAR_TEMP
      Index : Int;
   END_VAR
BEGIN

   #Cursor.Position := 0;
   #Cursor.First := 0;
   #Page.Revision := #Revision;
   #Page.PageIndex := 0;
   IF #PageIndex >= 0 AND #PageIndex <= 32767 THEN
       #Cursor.First := #PageIndex * 16;
       #Page.PageIndex := DINT_TO_INT(#PageIndex);
   END_IF;
   #Page.PageCount := 1;
   #Page.EntryCount := 0;
   "FRK_UnitScratch".EmptyConfigEntry.ValueType := 1;
   "FRK_UnitScratch".EmptyConfigEntry.Readable := TRUE;
   FOR #Index := 1 TO 16 DO
       #Page.Entries[#Index] := "FRK_UnitScratch".EmptyConfigEntry;
   END_FOR;
END_FUNCTION

FUNCTION "FRK_ConfigCatalog" : Void   // FC24, SCL
{ S7_Optimized_Access := 'TRUE' }
VERSION : 0.1
// stored: AutoNumber true, IsIECCheckEnabled false, SetENOAutomatically false, UDAEnableTagReadback false
   VAR_INPUT
      Scope : String;
      Count : Int;
      Catalog : Array[1..12] of "ST_CommandInfo";
      ReadLevel : DInt;
      Readable : Bool;
   END_VAR
   VAR_IN_OUT
      Cursor : "FRK_ConfigCursor";
      Page : "ST_ConfigPage";
   END_VAR
   VAR_TEMP
      Index : Int;
      IndexText : String[8];
      Prefix : String[254];
      Item : String[254];
   END_VAR
BEGIN

   "FRK_ConfigAppend"(Scope := #Scope,
                      Item := 'CatalogCount',
                      ValueText := STRING_TO_WSTRING(INT_TO_STRING(#Count)),
                      ValueType := 0,
                      ReadLevel := #ReadLevel,
                      Readable := #Readable,
                      Cursor := #Cursor,
                      Page := #Page);
   FOR #Index := 1 TO #Count DO
       IF #Index > 12 THEN
           EXIT;
       END_IF;
       #IndexText := INT_TO_STRING(#Index);
       IF #IndexText[1] = '+' THEN
           #IndexText := DELETE(IN := #IndexText, L := 1, P := 1);
       END_IF;
       #Prefix := CONCAT(IN1 := 'Catalog/Catalog[', IN2 := #IndexText);
       #Prefix := CONCAT(IN1 := #Prefix, IN2 := ']/');
       #Item := CONCAT(IN1 := #Prefix, IN2 := 'Value');
       "FRK_ConfigAppend"(Scope := #Scope,
                          Item := #Item,
                          ValueText := STRING_TO_WSTRING(DINT_TO_STRING(#Catalog[#Index].Value)),
                          ValueType := 0,
                          ReadLevel := #ReadLevel,
                          Readable := #Readable,
                          Cursor := #Cursor,
                          Page := #Page);
       #Item := CONCAT(IN1 := #Prefix, IN2 := 'Label');
       "FRK_ConfigAppend"(Scope := #Scope,
                          Item := #Item,
                          ValueText := STRING_TO_WSTRING(#Catalog[#Index].Label),
                          ValueType := 1,
                          ReadLevel := #ReadLevel,
                          Readable := #Readable,
                          Cursor := #Cursor,
                          Page := #Page);
       #Item := CONCAT(IN1 := #Prefix, IN2 := 'Style');
       "FRK_ConfigAppend"(Scope := #Scope,
                          Item := #Item,
                          ValueText := STRING_TO_WSTRING(DINT_TO_STRING(#Catalog[#Index].Style)),
                          ValueType := 0,
                          ReadLevel := #ReadLevel,
                          Readable := #Readable,
                          Cursor := #Cursor,
                          Page := #Page);
   END_FOR;
END_FUNCTION

FUNCTION "FRK_ConfigFinish" : Void   // FC23, SCL
{ S7_Optimized_Access := 'TRUE' }
VERSION : 0.1
// stored: AutoNumber true, IsIECCheckEnabled false, SetENOAutomatically false, UDAEnableTagReadback false
   VAR_IN_OUT
      Cursor : "FRK_ConfigCursor";
      Page : "ST_ConfigPage";
   END_VAR
BEGIN

   #Page.PageCount := DINT_TO_INT((#Cursor.Position + 16 - 1) / 16);
   IF #Page.PageCount < 1 THEN
       #Page.PageCount := 1;
   END_IF;
END_FUNCTION

FUNCTION "FRK_ConfigRevision" : UDInt   // FC20, SCL
{ S7_Optimized_Access := 'TRUE' }
VERSION : 0.1
// Core 3.10.2: deterministic typed walk, one bounded response window.
//  Static facets carry no write capability. Every reused slot is cleared.
// stored: AutoNumber true, IsIECCheckEnabled false, SetENOAutomatically false, UDAEnableTagReadback false
   VAR_INPUT
      Previous : UDInt;
   END_VAR
   VAR_TEMP
      Stamp : DTL;
      ResultCode : Int;
      Generation : ULInt;
   END_VAR
BEGIN

   #FRK_ConfigRevision := #Previous + 1;
   #ResultCode := RD_SYS_T(OUT => #Stamp);
   IF #ResultCode = 0 THEN
       #Generation := LDT_TO_ULINT(DTL_TO_LDT(#Stamp)) / ULINT#1000000;
       #FRK_ConfigRevision := ULINT_TO_UDINT(#Generation MOD ULINT#4294967296);
   END_IF;
   IF #FRK_ConfigRevision = #Previous THEN
       #FRK_ConfigRevision := #Previous + 1;
   END_IF;
   IF #FRK_ConfigRevision = 0 THEN
       #FRK_ConfigRevision := 1;
   END_IF;
END_FUNCTION

FUNCTION "FRK_ConfigUnit" : Void   // FC25, SCL
{ S7_Optimized_Access := 'TRUE' }
VERSION : 0.1
// stored: AutoNumber true, IsIECCheckEnabled false, SetENOAutomatically false, UDAEnableTagReadback false
   VAR_INPUT
      Scope : String;
      Policy : Array[0..6] of "ST_ModePolicy";
      ReadLevel : DInt;
      Readable : Bool;
   END_VAR
   VAR_IN_OUT
      Cursor : "FRK_ConfigCursor";
      Page : "ST_ConfigPage";
   END_VAR
   VAR_TEMP
      Index : Int;
      IndexText : String[8];
      Prefix : String[254];
      Item : String[254];
   END_VAR
BEGIN

   "FRK_ConfigAppend"(Scope := #Scope,
                      Item := 'CatalogCount',
                      ValueText := WSTRING#'0',
                      ValueType := 0,
                      ReadLevel := #ReadLevel,
                      Readable := #Readable,
                      Cursor := #Cursor,
                      Page := #Page);
   "FRK_ConfigAppend"(Scope := #Scope,
                      Item := 'AvailableModelCount',
                      ValueText := WSTRING#'0',
                      ValueType := 0,
                      ReadLevel := #ReadLevel,
                      Readable := #Readable,
                      Cursor := #Cursor,
                      Page := #Page);
   FOR #Index := 0 TO 6 DO
       #IndexText := INT_TO_STRING(#Index);
       IF #IndexText[1] = '+' THEN
           #IndexText := DELETE(IN := #IndexText, L := 1, P := 1);
       END_IF;
       #Prefix := CONCAT(IN1 := 'ModePolicy/ModePolicy[', IN2 := #IndexText);
       #Prefix := CONCAT(IN1 := #Prefix, IN2 := ']/');
       #Item := CONCAT(IN1 := #Prefix, IN2 := 'Shield');
       "FRK_ConfigAppend"(Scope := #Scope,
                          Item := #Item,
                          ValueText := STRING_TO_WSTRING(DINT_TO_STRING(#Policy[#Index].Shield)),
                          ValueType := 0,
                          ReadLevel := #ReadLevel,
                          Readable := #Readable,
                          Cursor := #Cursor,
                          Page := #Page);
       #Item := CONCAT(IN1 := #Prefix, IN2 := 'Style');
       "FRK_ConfigAppend"(Scope := #Scope,
                          Item := #Item,
                          ValueText := STRING_TO_WSTRING(DINT_TO_STRING(#Policy[#Index].Style)),
                          ValueType := 0,
                          ReadLevel := #ReadLevel,
                          Readable := #Readable,
                          Cursor := #Cursor,
                          Page := #Page);
   END_FOR;
END_FUNCTION

FUNCTION "FRK_Config_DeclarationCell" : Void   // FC64, SCL
{ S7_Optimized_Access := 'TRUE' }
VERSION : 0.1
// stored: AutoNumber true, IsIECCheckEnabled false, SetENOAutomatically false, UDAEnableTagReadback false
   VAR_INPUT
      ReadLevel : DInt;
      Readable : Bool;
   END_VAR
   VAR_IN_OUT
      Module : "FB_DeclarationCell";
      Cursor : "FRK_ConfigCursor";
      Page : "ST_ConfigPage";
   END_VAR
BEGIN

   "FRK_ConfigCatalog"(Scope := #Module.Status.Name,
                       Catalog := #Module.Catalog,
                       Count := #Module.CatalogCount,
                       ReadLevel := #ReadLevel,
                       Readable := #Readable,
                       Cursor := #Cursor,
                       Page := #Page);
   "FRK_Config_DeclarationCylinder"(Module := #Module.Clamp,
                                    ReadLevel := #ReadLevel,
                                    Readable := #Readable,
                                    Cursor := #Cursor,
                                    Page := #Page);
   "FRK_Config_DeclarationCylinder"(Module := #Module.Gate,
                                    ReadLevel := #ReadLevel,
                                    Readable := #Readable,
                                    Cursor := #Cursor,
                                    Page := #Page);
END_FUNCTION

FUNCTION "FRK_Config_DeclarationCylinder" : Void   // FC62, SCL
{ S7_Optimized_Access := 'TRUE' }
VERSION : 0.1
// stored: AutoNumber true, IsIECCheckEnabled false, SetENOAutomatically false, UDAEnableTagReadback false
   VAR_INPUT
      ReadLevel : DInt;
      Readable : Bool;
   END_VAR
   VAR_IN_OUT
      Module : "FB_DeclarationCylinder";
      Cursor : "FRK_ConfigCursor";
      Page : "ST_ConfigPage";
   END_VAR
BEGIN

   "FRK_ConfigCatalog"(Scope := #Module.Status.Name,
                       Catalog := #Module.Catalog,
                       Count := #Module.CatalogCount,
                       ReadLevel := #ReadLevel,
                       Readable := #Readable,
                       Cursor := #Cursor,
                       Page := #Page);
END_FUNCTION

FUNCTION "FRK_Config_DeclarationUnit" : Void   // FC73, SCL
{ S7_Optimized_Access := 'TRUE' }
VERSION : 0.1
// stored: AutoNumber true, IsIECCheckEnabled false, SetENOAutomatically false, UDAEnableTagReadback false
   VAR_INPUT
      ReadLevel : DInt;
      Readable : Bool;
   END_VAR
   VAR_IN_OUT
      Module : "FB_DeclarationUnit";
      Cursor : "FRK_ConfigCursor";
      Page : "ST_ConfigPage";
   END_VAR
BEGIN

   "FRK_ConfigUnit"(Scope := #Module.Status.Name,
                    Policy := #Module.ModePolicy,
                    ReadLevel := #ReadLevel,
                    Readable := #Readable,
                    Cursor := #Cursor,
                    Page := #Page);
   "FRK_Config_DeclarationCell"(Module := #Module.Cell,
                                ReadLevel := #ReadLevel,
                                Readable := #Readable,
                                Cursor := #Cursor,
                                Page := #Page);
   "FRK_Config_SatelliteUnit"(Module := #Module.Satellite,
                              ReadLevel := #ReadLevel,
                              Readable := #Readable,
                              Cursor := #Cursor,
                              Page := #Page);
END_FUNCTION

FUNCTION "FRK_Config_InnerUnit" : Void   // FC67, SCL
{ S7_Optimized_Access := 'TRUE' }
VERSION : 0.1
// stored: AutoNumber true, IsIECCheckEnabled false, SetENOAutomatically false, UDAEnableTagReadback false
   VAR_INPUT
      ReadLevel : DInt;
      Readable : Bool;
   END_VAR
   VAR_IN_OUT
      Module : "FB_InnerUnit";
      Cursor : "FRK_ConfigCursor";
      Page : "ST_ConfigPage";
   END_VAR
BEGIN

   "FRK_ConfigUnit"(Scope := #Module.Status.Name,
                    Policy := #Module.ModePolicy,
                    ReadLevel := #ReadLevel,
                    Readable := #Readable,
                    Cursor := #Cursor,
                    Page := #Page);
   "FRK_Config_DeclarationCell"(Module := #Module.Cell,
                                ReadLevel := #ReadLevel,
                                Readable := #Readable,
                                Cursor := #Cursor,
                                Page := #Page);
END_FUNCTION

FUNCTION "FRK_Config_SatelliteUnit" : Void   // FC70, SCL
{ S7_Optimized_Access := 'TRUE' }
VERSION : 0.1
// stored: AutoNumber true, IsIECCheckEnabled false, SetENOAutomatically false, UDAEnableTagReadback false
   VAR_INPUT
      ReadLevel : DInt;
      Readable : Bool;
   END_VAR
   VAR_IN_OUT
      Module : "FB_SatelliteUnit";
      Cursor : "FRK_ConfigCursor";
      Page : "ST_ConfigPage";
   END_VAR
BEGIN

   "FRK_ConfigUnit"(Scope := #Module.Status.Name,
                    Policy := #Module.ModePolicy,
                    ReadLevel := #ReadLevel,
                    Readable := #Readable,
                    Cursor := #Cursor,
                    Page := #Page);
   "FRK_Config_DeclarationCell"(Module := #Module.Cell,
                                ReadLevel := #ReadLevel,
                                Readable := #Readable,
                                Cursor := #Cursor,
                                Page := #Page);
   "FRK_Config_InnerUnit"(Module := #Module.Inner,
                          ReadLevel := #ReadLevel,
                          Readable := #Readable,
                          Cursor := #Cursor,
                          Page := #Page);
END_FUNCTION

FUNCTION "FRK_DescendantsReady" : Bool   // FC50, SCL
{ S7_Optimized_Access := 'TRUE' }
VERSION : 0.1
// stored: AutoNumber true, IsIECCheckEnabled false, SetENOAutomatically false, UDAEnableTagReadback false
   VAR_INPUT
      OwnerIndex : DInt;
   END_VAR
   VAR_TEMP
      Index : DInt;
      Parent : DInt;
      Depth : DInt;
   END_VAR
BEGIN

   #FRK_DescendantsReady := FALSE;
   IF "FRK_Registry".Fault OR #OwnerIndex < 1 OR #OwnerIndex > "FRK_Registry".Count OR "FRK_Registry".Count > 32 THEN
       RETURN;
   END_IF;
   FOR #Index := 1 TO "FRK_Registry".Count DO
       #Parent := "FRK_Registry".Rows[#Index].Parent;
       FOR #Depth := 1 TO 32 DO
           IF #Parent = #OwnerIndex THEN
               IF "FRK_Registry".Rows[#Index].Exec <> 0 THEN
                   RETURN;
               END_IF;
               EXIT;
           END_IF;
           IF #Parent = 0 THEN
               EXIT;
           END_IF;
           IF #Parent < 1 OR #Parent > "FRK_Registry".Count THEN
               RETURN;
           END_IF;
           #Parent := "FRK_Registry".Rows[#Parent].Parent;
       END_FOR;
       IF #Depth > 32 AND #Parent <> 0 THEN
           RETURN;
       END_IF;
   END_FOR;
   #FRK_DescendantsReady := TRUE;
END_FUNCTION

FUNCTION "FRK_Diagnostic" : Void   // FC7, SCL
{ S7_Optimized_Access := 'TRUE' }
VERSION : 0.1
// stored: AutoNumber true, IsIECCheckEnabled false, SetENOAutomatically false, UDAEnableTagReadback false
   VAR_INPUT
      ReasonCode : DInt;
      Description : WString;
      Severity : DInt;
   END_VAR
   VAR_IN_OUT
      Status : "ST_ModuleStatus";
   END_VAR
   VAR_TEMP
      Stamp : DTL;
      ResultCode : Int;
   END_VAR
BEGIN

   #Status.Diagnostic.ReasonCode := #ReasonCode;
   #Status.Diagnostic.SourcePath := STRING_TO_WSTRING(#Status.Name);
   #Status.Diagnostic.Description := #Description;
   #Status.Diagnostic.IoTag := '';
   #Status.Diagnostic.IoAddress := '';
   #Status.Diagnostic.Severity := #Severity;
   #Status.Diagnostic.Category := 0;
   #ResultCode := RD_SYS_T(OUT => #Stamp);
   IF #ResultCode = 0 THEN
       #Status.Diagnostic.Since := DTL_TO_LDT(#Stamp);
   ELSE
       #Status.Diagnostic.Since := LDT#1970-01-01-00:00:00.000000000;
   END_IF;
   // UTC source alone is not proof of synchronization; quality stays false.
   #Status.Diagnostic.TimeSynchronized := FALSE;
END_FUNCTION

FUNCTION "FRK_Elapsed" : UDInt   // FC4, SCL
{ S7_Optimized_Access := 'TRUE' }
VERSION : 0.1
// stored: AutoNumber true, IsIECCheckEnabled false, SetENOAutomatically false, UDAEnableTagReadback false
   VAR_INPUT
      NewMs : UDInt;
      OldMs : UDInt;
   END_VAR
   VAR_TEMP
      Wide : ULInt;
   END_VAR
BEGIN

   IF #NewMs >= #OldMs THEN
       #Wide := UDINT_TO_ULINT(#NewMs) - UDINT_TO_ULINT(#OldMs);
   ELSE
       #Wide := ULINT#4294967296 + UDINT_TO_ULINT(#NewMs) - UDINT_TO_ULINT(#OldMs);
   END_IF;
   #FRK_Elapsed := ULINT_TO_UDINT(#Wide);
END_FUNCTION

FUNCTION "FRK_End" : Void   // FC18, SCL
{ S7_Optimized_Access := 'TRUE' }
VERSION : 0.1
// stored: AutoNumber true, IsIECCheckEnabled false, SetENOAutomatically false, UDAEnableTagReadback false
   VAR_OUTPUT
      Busy : Bool;
      Done : Bool;
      Error : Bool;
      Aborted : Bool;
      Held : Bool;
      ErrorID : DWord;
      Timing : "ST_ModuleTiming";
   END_VAR
   VAR_IN_OUT
      Core : "FRK_Core";
      Status : "ST_ModuleStatus";
   END_VAR
   VAR_TEMP
      ActiveWide : ULInt;
   END_VAR
BEGIN

   IF #Core.Exec = 1 THEN
       IF #Core.Held AND NOT #Core.HoldReq AND NOT #Core.DiagTouched THEN
           "FRK_ClearDiag"(Status := #Status);
       END_IF;
       // HELD suspends progress timeout. Wall-clock command duration includes it.
       IF NOT #Core.Held AND NOT #Core.HoldReq THEN
           #ActiveWide := UDINT_TO_ULINT(#Core.ActiveMs) + UDINT_TO_ULINT(#Core.DeltaMs);
           IF #ActiveWide > ULINT#2147483647 THEN
               #ActiveWide := ULINT#2147483647;
           END_IF;
           #Core.ActiveMs := ULINT_TO_UDINT(#ActiveWide);
           IF #Core.TimeoutMs > 0 AND #Core.ActiveMs >= #Core.TimeoutMs THEN
               IF #Status.Diagnostic.ReasonCode = 0 THEN
                   "FRK_Fault"(Core := #Core,
                               Status := #Status,
                               ReasonCode := 2001,
                               Description := WSTRING#'fraktal.command.timeout');
               ELSE
                   #Status.Diagnostic.Severity := 1;
                   "FRK_Rationalize"(Diag := #Status.Diagnostic);
                   #Core.Exec := 3;
                   #Core.Step := 0;
                   #Core.Dispatch := FALSE;
               END_IF;
           END_IF;
       END_IF;
   END_IF;
   #Core.Held := #Core.HoldReq AND #Core.Exec = 1;
   IF NOT #Core.Held THEN
       #Core.HoldReason := 0;
   END_IF;
   IF #Core.TimingOpen AND #Core.Exec <> 1 THEN
       "FRK_RecordTiming"(Core := #Core);
   END_IF;
   #Busy := #Core.Exec = 1;
   #Done := #Core.Exec = 2;
   #Error := #Core.Exec = 3;
   #Aborted := #Core.Exec = 4;
   #Held := #Core.Held;
   #ErrorID := DINT_TO_DWORD(#Status.Diagnostic.ReasonCode);
   #Timing := #Core.Timing;
   #Status.State := #Core.Exec;
   #Status.FaultActive := #Core.Exec = 3;
   #Core.HoldReq := FALSE;
   #Core.EvInit := FALSE;
   #Core.EvCommandStart := FALSE;
   #Core.EvAbort := FALSE;
   #Core.EvAbortInError := FALSE;
   #Core.ReleasePending := FALSE;
   "FRK_SyncRegistry"(Index := #Core.RegIndex,
                      Status := #Status);
END_FUNCTION

FUNCTION "FRK_Fault" : Void   // FC8, SCL
{ S7_Optimized_Access := 'TRUE' }
VERSION : 0.1
// stored: AutoNumber true, IsIECCheckEnabled false, SetENOAutomatically false, UDAEnableTagReadback false
   VAR_INPUT
      ReasonCode : DInt;
      Description : WString;
   END_VAR
   VAR_IN_OUT
      Core : "FRK_Core";
      Status : "ST_ModuleStatus";
   END_VAR
BEGIN

   IF #Core.Exec = 3 THEN
       RETURN;
   END_IF;
   "FRK_Diagnostic"(Status := #Status,
                    ReasonCode := #ReasonCode,
                    Description := #Description,
                    Severity := 1);
   "FRK_Rationalize"(Diag := #Status.Diagnostic);
   #Core.Exec := 3;
   #Core.Step := 0;
   #Core.Dispatch := FALSE;
   #Core.DiagTouched := TRUE;
END_FUNCTION

FUNCTION "FRK_HistoryEvent" : Void   // FC52, SCL
{ S7_Optimized_Access := 'TRUE' }
VERSION : 0.1
// Shared Unit routing: typed generated edges carry these owning predicates.
// stored: AutoNumber true, IsIECCheckEnabled false, SetENOAutomatically false, UDAEnableTagReadback false
   VAR_INPUT
      Reason : DInt;
      Description : WString;
      SourcePath : WString;
   END_VAR
   VAR_IN_OUT
      History : Array[1..16] of "ST_Diagnostic";
      Head : Int;
   END_VAR
   VAR_TEMP
      Stamp : DTL;
      ResultCode : Int;
   END_VAR
BEGIN

   IF #Head < 0 OR #Head >= 16 THEN
       #Head := 0;
   END_IF;
   #Head := #Head + 1;
   #History[#Head] := "FRK_UnitScratch".EmptyDiagnostic;
   #History[#Head].ReasonCode := #Reason;
   #History[#Head].Description := #Description;
   #History[#Head].SourcePath := #SourcePath;
   #History[#Head].Severity := 0;
   #History[#Head].Category := 2;
   #ResultCode := RD_SYS_T(OUT => #Stamp);
   IF #ResultCode = 0 THEN
       #History[#Head].Since := DTL_TO_LDT(#Stamp);
   END_IF;
END_FUNCTION

FUNCTION "FRK_Hold" : Void   // FC11, SCL
{ S7_Optimized_Access := 'TRUE' }
VERSION : 0.1
// stored: AutoNumber true, IsIECCheckEnabled false, SetENOAutomatically false, UDAEnableTagReadback false
   VAR_INPUT
      ReasonCode : DInt;
      Description : WString;
   END_VAR
   VAR_IN_OUT
      Core : "FRK_Core";
      Status : "ST_ModuleStatus";
   END_VAR
BEGIN

   IF #Core.Exec <> 1 THEN
       RETURN;
   END_IF;
   IF NOT #Core.Held OR #Core.HoldReason <> #ReasonCode THEN
       "FRK_Diagnostic"(Status := #Status,
                        ReasonCode := #ReasonCode,
                        Description := #Description,
                        Severity := 0);
   END_IF;
   #Core.HoldReq := TRUE;
   #Core.HoldReason := #ReasonCode;
   #Core.DiagTouched := TRUE;
END_FUNCTION

FUNCTION "FRK_HoldDiag" : Void   // FC10, SCL
{ S7_Optimized_Access := 'TRUE' }
VERSION : 0.1
// stored: AutoNumber true, IsIECCheckEnabled false, SetENOAutomatically false, UDAEnableTagReadback false
   VAR_INPUT
      Diag : "ST_Diagnostic";
   END_VAR
   VAR_IN_OUT
      Core : "FRK_Core";
      Status : "ST_ModuleStatus";
   END_VAR
BEGIN

   IF #Core.Exec <> 1 THEN
       RETURN;
   END_IF;
   #Status.Diagnostic := #Diag;
   #Status.Diagnostic.Severity := 0;
   #Core.HoldReq := TRUE;
   #Core.HoldReason := #Diag.ReasonCode;
   #Core.DiagTouched := TRUE;
END_FUNCTION

FUNCTION "FRK_ManualApply" : Void   // FC57, SCL
{ S7_Optimized_Access := 'TRUE' }
VERSION : 0.1
// stored: AutoNumber true, IsIECCheckEnabled false, SetENOAutomatically false, UDAEnableTagReadback false
   VAR_INPUT
      Request : "ST_HmiRequest";
      Status : "ST_ModuleStatus";
      Core : "FRK_Core";
      Commands : Array[1..12] of "ST_CommandInfo";
      Count : DInt;
      Conditions : Array[1..16] of "FRK_ManualConditionRow";
   END_VAR
   VAR_IN_OUT
      Report : "ST_ReleaseReport";
      Execute : Bool;
      Command : DInt;
      ManualOwned : Bool;
   END_VAR
   VAR_TEMP
      Index : Int;
      Supported : Bool;
      PreviousCount : Int;
   END_VAR
BEGIN

   #Supported := FALSE;
   IF #Count >= 0 AND #Count <= 12 THEN
       FOR #Index := 1 TO DINT_TO_INT(#Count) DO
           IF #Commands[#Index].Value = #Request.IntValue AND #Commands[#Index].Style = 0 THEN
               #Supported := TRUE;
           END_IF;
       END_FOR;
   END_IF;
   IF NOT #Supported THEN
       "FRK_ReleaseReason"(Report := #Report,
                           Description := WSTRING#'std.error.unsupportedHmiRequest',
                           Reason := 2008,
                           Path := STRING_TO_WSTRING(#Status.Name),
                           Kind := 4);
   END_IF;
   IF #Core.Exec <> 0 OR #Execute OR #Core.ReleasePending THEN
       "FRK_ReleaseReason"(Report := #Report,
                           Description := WSTRING#'std.error.hmiRequestRejected',
                           Reason := 2011,
                           Path := STRING_TO_WSTRING(#Status.Name),
                           Kind := 4);
   END_IF;
   FOR #Index := 1 TO 16 DO
       IF #Conditions[#Index].Used AND NOT #Conditions[#Index].Ok THEN
           IF #Conditions[#Index].Value = 0 OR #Conditions[#Index].Value = #Request.IntValue THEN
               #PreviousCount := #Report.Count;
               "FRK_ReleaseReason"(Report := #Report,
                                   Description := #Conditions[#Index].Diag.Description,
                                   Reason := #Conditions[#Index].Diag.ReasonCode,
                                   Path := STRING_TO_WSTRING(#Status.Name),
                                   Kind := 3);
               IF #Report.Count > #PreviousCount THEN
                   #Report.Reasons[#Report.Count].Bypassable := #Conditions[#Index].Bypassable;
               END_IF;
           END_IF;
       END_IF;
   END_FOR;
   IF #Request.Kind = 11 AND #Report.Released THEN
       #Command := #Request.IntValue;
       #Execute := TRUE;
       #ManualOwned := TRUE;
   END_IF;
END_FUNCTION

FUNCTION "FRK_ManualCommon" : Void   // FC55, SCL
{ S7_Optimized_Access := 'TRUE' }
VERSION : 0.1
// stored: AutoNumber true, IsIECCheckEnabled false, SetENOAutomatically false, UDAEnableTagReadback false
   VAR_INPUT
      Core : "FRK_Core";
      Unit : "FRK_Unit";
      Status : "ST_ModuleStatus";
   END_VAR
   VAR_IN_OUT
      Report : "ST_ReleaseReport";
   END_VAR
BEGIN

   IF #Unit.Mode <> 1 OR #Unit.ModePending THEN
       "FRK_ReleaseReason"(Report := #Report,
                           Description := WSTRING#'std.release.manualModeRequired',
                           Reason := 2002,
                           Path := STRING_TO_WSTRING(#Status.Name),
                           Kind := 0);
   END_IF;
   IF #Core.Exec <> 0 OR #Unit.Clearing OR #Unit.FaultLatched THEN
       "FRK_ReleaseReason"(Report := #Report,
                           Description := WSTRING#'std.error.hmiRequestRejected',
                           Reason := 2011,
                           Path := STRING_TO_WSTRING(#Status.Name),
                           Kind := 4);
   END_IF;
   IF NOT #Unit.Permit THEN
       "FRK_ReleaseReason"(Report := #Report,
                           Description := #Unit.PermitDiag.Description,
                           Reason := #Unit.PermitDiag.ReasonCode,
                           Path := #Unit.PermitDiag.SourcePath,
                           Kind := 3);
   END_IF;
END_FUNCTION

FUNCTION "FRK_ManualCondition" : Void   // FC56, SCL
{ S7_Optimized_Access := 'TRUE' }
VERSION : 0.1
// stored: AutoNumber true, IsIECCheckEnabled false, SetENOAutomatically false, UDAEnableTagReadback false
   VAR_INPUT
      Slot : Int;
      Value : DInt;
      Ok : Bool;
      Diag : "ST_Diagnostic";
      Bypassable : Bool;
   END_VAR
   VAR_IN_OUT
      Conditions : Array[1..16] of "FRK_ManualConditionRow";
   END_VAR
BEGIN

   IF #Slot < 1 OR #Slot > 16 THEN
       RETURN;
   END_IF;
   #Conditions[#Slot].Used := TRUE;
   #Conditions[#Slot].Value := #Value;
   #Conditions[#Slot].Ok := #Ok;
   #Conditions[#Slot].Diag := #Diag;
   #Conditions[#Slot].Bypassable := #Bypassable;
END_FUNCTION

FUNCTION "FRK_ManualFinish" : Void   // FC58, SCL
{ S7_Optimized_Access := 'TRUE' }
VERSION : 0.1
// stored: AutoNumber true, IsIECCheckEnabled false, SetENOAutomatically false, UDAEnableTagReadback false
   VAR_INPUT
      Core : "FRK_Core";
   END_VAR
   VAR_IN_OUT
      Execute : Bool;
      ManualOwned : Bool;
   END_VAR
BEGIN

   IF #ManualOwned AND #Core.Exec <> 1 THEN
       #Execute := FALSE;
       #ManualOwned := FALSE;
   END_IF;
END_FUNCTION

FUNCTION "FRK_PartAborted" : Void   // FC41, SCL
{ S7_Optimized_Access := 'TRUE' }
VERSION : 0.1
// stored: AutoNumber true, IsIECCheckEnabled false, SetENOAutomatically false, UDAEnableTagReadback false
   VAR_IN_OUT
      Core : "FRK_Core";
      Unit : "FRK_Unit";
      Status : "ST_ModuleStatus";
      Part : "ST_PartContext";
      History : Array[1..16] of "ST_Diagnostic";
      Head : Int;
   END_VAR
BEGIN

   IF #Unit.CarrierIndex = 0 OR NOT #Part.Present THEN
       RETURN;
   END_IF;
   #Part.Result.Verdict := 0;
   IF #Core.Exec = 3 AND #Part.Result.ReasonCode = 0 THEN
       #Part.Result.ReasonCode := #Status.Diagnostic.ReasonCode;
   END_IF;
   "FRK_PartEvent"(History := #History,
                   Head := #Head,
                   Reason := 2027,
                   Uid := #Part.Uid,
                   SourcePath := #Status.Name);
   #Part.Present := FALSE;
END_FUNCTION

FUNCTION "FRK_PartEvent" : Void   // FC37, SCL
{ S7_Optimized_Access := 'TRUE' }
VERSION : 0.1
// stored: AutoNumber true, IsIECCheckEnabled false, SetENOAutomatically false, UDAEnableTagReadback false
   VAR_INPUT
      Reason : DInt;
      Uid : String;
      SourcePath : String;
   END_VAR
   VAR_IN_OUT
      History : Array[1..16] of "ST_Diagnostic";
      Head : Int;
   END_VAR
   VAR_TEMP
      Stamp : DTL;
      ResultCode : Int;
   END_VAR
BEGIN

   IF #Head < 0 OR #Head >= 16 THEN
       #Head := 0;
   END_IF;
   #Head := #Head + 1;
   #History[#Head].ReasonCode := #Reason;
   #History[#Head].SourcePath := STRING_TO_WSTRING(#SourcePath);
   CASE #Reason OF
       2024:
           #History[#Head].Description := WSTRING#'std.event.partReceived: ';
       2025:
           #History[#Head].Description := WSTRING#'std.event.partProcessingStarted: ';
       2026:
           #History[#Head].Description := WSTRING#'std.event.partProcessed: ';
       2027:
           #History[#Head].Description := WSTRING#'std.event.partAborted: ';
       ELSE
           #History[#Head].Description := WSTRING#'';
   END_CASE;
   #History[#Head].Description := CONCAT(IN1 := #History[#Head].Description, IN2 := STRING_TO_WSTRING(#Uid));
   #History[#Head].IoTag := '';
   #History[#Head].IoAddress := '';
   #History[#Head].Severity := 0;
   #History[#Head].Category := 0;
   #History[#Head].TimeSynchronized := FALSE;
   #History[#Head].Since := LDT#1970-01-01-00:00:00.000000000;
   #ResultCode := RD_SYS_T(OUT => #Stamp);
   IF #ResultCode = 0 THEN
       #History[#Head].Since := DTL_TO_LDT(#Stamp);
   END_IF;
END_FUNCTION

FUNCTION "FRK_PartProcessed" : Bool   // FC40, SCL
{ S7_Optimized_Access := 'TRUE' }
VERSION : 0.1
// stored: AutoNumber true, IsIECCheckEnabled false, SetENOAutomatically false, UDAEnableTagReadback false
   VAR_INPUT
      Verdict : DInt;
      Reason : DInt;
   END_VAR
   VAR_IN_OUT
      Core : "FRK_Core";
      Unit : "FRK_Unit";
      Status : "ST_ModuleStatus";
      Part : "ST_PartContext";
      History : Array[1..16] of "ST_Diagnostic";
      Head : Int;
   END_VAR
   VAR_TEMP
      Index : DInt;
      Stamp : DTL;
      ResultCode : Int;
   END_VAR
BEGIN

   #FRK_PartProcessed := FALSE;
   #Index := #Unit.CarrierIndex;
   IF #Index = 0 OR NOT #Part.Present THEN
       RETURN;
   END_IF;
   IF #Verdict < 1 OR #Verdict > 3 OR (#Verdict = 2 AND #Reason = 0) THEN
       "FRK_Fault"(Core := #Core,
                   Status := #Status,
                   ReasonCode := 2023,
                   Description := WSTRING#'std.error.nokReasonRequired');
       RETURN;
   END_IF;
   IF #Index < 1 OR #Index > 32 THEN
       "FRK_Fault"(Core := #Core,
                   Status := #Status,
                   ReasonCode := 2021,
                   Description := WSTRING#'std.error.partCarrierWriteFailed');
       RETURN;
   END_IF;
   IF NOT "FRK_Carriers".Slots[#Index].Enabled THEN
       "FRK_Fault"(Core := #Core,
                   Status := #Status,
                   ReasonCode := 2021,
                   Description := WSTRING#'std.error.partCarrierWriteFailed');
       RETURN;
   END_IF;
   IF #Part.Uid <> "FRK_Carriers".Slots[#Index].Context.Uid THEN
       "FRK_Fault"(Core := #Core,
                   Status := #Status,
                   ReasonCode := 2022,
                   Description := WSTRING#'std.error.partCarrierReadFailed');
       RETURN;
   END_IF;
   #Part.Result.Verdict := #Verdict;
   #Part.Result.ReasonCode := #Reason;
   #Part.Result.StationPath := STRING_TO_WSTRING(#Status.Name);
   #Part.Result.TimeSynchronized := FALSE;
   #ResultCode := RD_SYS_T(OUT => #Stamp);
   IF #ResultCode = 0 THEN
       #Part.Result.Stamp := DTL_TO_LDT(#Stamp);
   END_IF;
   "FRK_Carriers".Slots[#Index].Written := #Part;
   IF "FRK_Carriers".Slots[#Index].Writes < UDINT#4294967295 THEN
       "FRK_Carriers".Slots[#Index].Writes := "FRK_Carriers".Slots[#Index].Writes + 1;
   END_IF;
   CASE #Verdict OF
       1:
           IF #Unit.Good < UDINT#4294967295 THEN
               #Unit.Good := #Unit.Good + 1;
           END_IF;
       2:
           IF #Unit.Nok < UDINT#4294967295 THEN
               #Unit.Nok := #Unit.Nok + 1;
           END_IF;
           #Unit.NokReason := #Reason;
       3:
           IF #Unit.Rework < UDINT#4294967295 THEN
               #Unit.Rework := #Unit.Rework + 1;
           END_IF;
       ELSE
           RETURN;
   END_CASE;
   // The provider result is written before publishing EVENT_PART_PROCESSED.
   "FRK_PartEvent"(History := #History,
                   Head := #Head,
                   Reason := 2026,
                   Uid := #Part.Uid,
                   SourcePath := #Status.Name);
   #Part.Present := FALSE;
   #FRK_PartProcessed := TRUE;
END_FUNCTION

FUNCTION "FRK_PartReceived" : Bool   // FC38, SCL
{ S7_Optimized_Access := 'TRUE' }
VERSION : 0.1
// stored: AutoNumber true, IsIECCheckEnabled false, SetENOAutomatically false, UDAEnableTagReadback false
   VAR_IN_OUT
      Core : "FRK_Core";
      Unit : "FRK_Unit";
      Status : "ST_ModuleStatus";
      Part : "ST_PartContext";
      History : Array[1..16] of "ST_Diagnostic";
      Head : Int;
   END_VAR
   VAR_TEMP
      Index : DInt;
      Uid : String[64];
      ResultIndex : DInt;
   END_VAR
BEGIN

   #FRK_PartReceived := FALSE;
   #Index := #Unit.CarrierIndex;
   IF #Index = 0 THEN
       RETURN;
   END_IF;
   IF #Index < 1 OR #Index > 32 THEN
       "FRK_Fault"(Core := #Core,
                   Status := #Status,
                   ReasonCode := 2020,
                   Description := WSTRING#'std.error.partCarrierReadFailed');
       RETURN;
   END_IF;
   IF NOT "FRK_Carriers".Slots[#Index].Enabled OR "FRK_Carriers".Slots[#Index].Kind <> 2 OR "FRK_Carriers".Slots[#Index].Serial = UDINT#4294967295 THEN
       "FRK_Fault"(Core := #Core,
                   Status := #Status,
                   ReasonCode := 2020,
                   Description := WSTRING#'std.error.partCarrierReadFailed');
       RETURN;
   END_IF;
   "FRK_Carriers".Slots[#Index].Serial := "FRK_Carriers".Slots[#Index].Serial + 1;
   #Uid := CONCAT(IN1 := 'FRK-', IN2 := DINT_TO_STRING(#Index));
   #Uid := CONCAT(IN1 := #Uid, IN2 := '-');
   #Uid := CONCAT(IN1 := #Uid, IN2 := UDINT_TO_STRING("FRK_Carriers".Slots[#Index].Serial));
   #Part.Uid := #Uid;
   #Part.Present := TRUE;
   #Part.CarrierKind := 2;
   #Part.Result.Verdict := 0;
   #Part.Result.ReasonCode := 0;
   #Part.Result.StationPath := STRING_TO_WSTRING(#Status.Name);
   #Part.Result.Stamp := LDT#1970-01-01-00:00:00.000000000;
   #Part.Result.TimeSynchronized := FALSE;
   FOR #ResultIndex := 1 TO 32 DO
       #Part.Result.Records[#ResultIndex].Name := '';
   END_FOR;
   FOR #ResultIndex := 1 TO 8 DO
       #Part.Parents[#ResultIndex] := '';
   END_FOR;
   "FRK_Carriers".Slots[#Index].Context := #Part;
   "FRK_PartEvent"(History := #History,
                   Head := #Head,
                   Reason := 2024,
                   Uid := #Part.Uid,
                   SourcePath := #Status.Name);
   #FRK_PartReceived := TRUE;
END_FUNCTION

FUNCTION "FRK_PartStarted" : Void   // FC39, SCL
{ S7_Optimized_Access := 'TRUE' }
VERSION : 0.1
// stored: AutoNumber true, IsIECCheckEnabled false, SetENOAutomatically false, UDAEnableTagReadback false
   VAR_IN_OUT
      Unit : "FRK_Unit";
      Status : "ST_ModuleStatus";
      Part : "ST_PartContext";
      History : Array[1..16] of "ST_Diagnostic";
      Head : Int;
   END_VAR
BEGIN

   IF #Unit.CarrierIndex = 0 OR NOT #Part.Present THEN
       RETURN;
   END_IF;
   "FRK_PartEvent"(History := #History,
                   Head := #Head,
                   Reason := 2025,
                   Uid := #Part.Uid,
                   SourcePath := #Status.Name);
END_FUNCTION

FUNCTION "FRK_PathOwned" : Bool   // FC53, SCL
{ S7_Optimized_Access := 'TRUE' }
VERSION : 0.1
// stored: AutoNumber true, IsIECCheckEnabled false, SetENOAutomatically false, UDAEnableTagReadback false
   VAR_INPUT
      OwnerPath : String;
      TargetPath : WString;
   END_VAR
   VAR_TEMP
      Width : Int;
   END_VAR
BEGIN

   #FRK_PathOwned := FALSE;
   #Width := LEN(#OwnerPath);
   IF #Width = 0 THEN
       RETURN;
   END_IF;
   IF #TargetPath = STRING_TO_WSTRING(#OwnerPath) THEN
       #FRK_PathOwned := TRUE;
       RETURN;
   END_IF;
   IF LEN(#TargetPath) <= #Width THEN
       RETURN;
   END_IF;
   #FRK_PathOwned := LEFT(IN := #TargetPath, L := #Width) = STRING_TO_WSTRING(#OwnerPath) AND #TargetPath[#Width + 1] = WCHAR#'.';
END_FUNCTION

FUNCTION "FRK_Pending" : Void   // FC12, SCL
{ S7_Optimized_Access := 'TRUE' }
VERSION : 0.1
// stored: AutoNumber true, IsIECCheckEnabled false, SetENOAutomatically false, UDAEnableTagReadback false
   VAR_INPUT
      Diag : "ST_Diagnostic";
   END_VAR
   VAR_IN_OUT
      Core : "FRK_Core";
      Status : "ST_ModuleStatus";
   END_VAR
BEGIN

   IF #Core.Exec = 1 AND NOT #Core.DiagTouched THEN
       #Status.Diagnostic := #Diag;
       #Status.Diagnostic.Severity := 0;
       #Core.DiagTouched := TRUE;
   END_IF;
END_FUNCTION

FUNCTION "FRK_Rationalize" : Void   // FC6, SCL
{ S7_Optimized_Access := 'TRUE' }
VERSION : 0.1
// stored: AutoNumber true, IsIECCheckEnabled false, SetENOAutomatically false, UDAEnableTagReadback false
   VAR_IN_OUT
      Diag : "ST_Diagnostic";
   END_VAR
BEGIN

   CASE #Diag.ReasonCode OF
       10:
           #Diag.Severity := 1;
           #Diag.Category := 2;
       11:
           #Diag.Severity := 0;
           #Diag.Category := 2;
       12:
           #Diag.Severity := 0;
           #Diag.Category := 2;
       13:
           #Diag.Severity := 1;
           #Diag.Category := 2;
       14:
           #Diag.Severity := 1;
           #Diag.Category := 2;
       15:
           #Diag.Severity := 2;
           #Diag.Category := 2;
       16:
           #Diag.Severity := 0;
           #Diag.Category := 2;
       17:
           #Diag.Severity := 0;
           #Diag.Category := 2;
       18:
           #Diag.Severity := 1;
           #Diag.Category := 2;
       19:
           #Diag.Severity := 0;
           #Diag.Category := 2;
       20:
           #Diag.Severity := 1;
           #Diag.Category := 2;
       21:
           #Diag.Severity := 0;
           #Diag.Category := 2;
       2001:
           #Diag.Severity := 1;
           #Diag.Category := 0;
       2002:
           #Diag.Severity := 0;
           #Diag.Category := 0;
       2003:
           #Diag.Severity := 1;
           #Diag.Category := 0;
       2004:
           #Diag.Severity := 1;
           #Diag.Category := 0;
       2005:
           #Diag.Severity := 0;
           #Diag.Category := 0;
       2006:
           #Diag.Severity := 1;
           #Diag.Category := 0;
       2007:
           #Diag.Severity := 0;
           #Diag.Category := 0;
       2008:
           #Diag.Severity := 0;
           #Diag.Category := 0;
       2010:
           #Diag.Severity := 1;
           #Diag.Category := 2;
       2011:
           #Diag.Severity := 0;
           #Diag.Category := 0;
       2012:
           #Diag.Severity := 1;
           #Diag.Category := 2;
       2020:
           #Diag.Severity := 1;
           #Diag.Category := 2;
       2021:
           #Diag.Severity := 1;
           #Diag.Category := 2;
       2022:
           #Diag.Severity := 2;
           #Diag.Category := 0;
       2023:
           #Diag.Severity := 1;
           #Diag.Category := 0;
       2024:
           #Diag.Severity := 0;
           #Diag.Category := 0;
       2025:
           #Diag.Severity := 0;
           #Diag.Category := 0;
       2026:
           #Diag.Severity := 0;
           #Diag.Category := 0;
       2027:
           #Diag.Severity := 0;
           #Diag.Category := 0;
       2030:
           #Diag.Severity := 0;
           #Diag.Category := 2;
       2040:
           #Diag.Severity := 1;
           #Diag.Category := 2;
       2041:
           #Diag.Severity := 1;
           #Diag.Category := 2;
       2042:
           #Diag.Severity := 0;
           #Diag.Category := 2;
       2043:
           #Diag.Severity := 0;
           #Diag.Category := 2;
       2901:
           #Diag.Severity := 0;
           #Diag.Category := 2;
       ELSE
           RETURN;
   END_CASE;
END_FUNCTION

FUNCTION "FRK_RecordTiming" : Void   // FC17, SCL
{ S7_Optimized_Access := 'TRUE' }
VERSION : 0.1
// stored: AutoNumber true, IsIECCheckEnabled false, SetENOAutomatically false, UDAEnableTagReadback false
   VAR_IN_OUT
      Core : "FRK_Core";
   END_VAR
   VAR_TEMP
      Index : DInt;
      Slot : DInt;
      DurationMs : UDInt;
      AverageMs : LInt;
   END_VAR
BEGIN

   #DurationMs := "FRK_Elapsed"(NewMs := "FRK_Clock".NowMs, OldMs := #Core.StartMs);
   // TIME's positive domain is bounded; clamp instead of publishing negatives.
   IF #DurationMs > UDINT#2147483647 THEN
       #DurationMs := UDINT#2147483647;
   END_IF;
   #Core.Timing.LastCmdTime := DINT_TO_TIME(UDINT_TO_DINT(#DurationMs));
   #Slot := 0;
   FOR #Index := 1 TO 8 DO
       IF #Core.Timing.Rows[#Index].Count > 0 AND #Core.Timing.Rows[#Index].Id = #Core.Command THEN
           #Slot := #Index;
           EXIT;
       ELSIF #Slot = 0 AND #Core.Timing.Rows[#Index].Count = 0 THEN
           #Slot := #Index;
       END_IF;
   END_FOR;
   IF #Slot = 0 THEN
       #Core.Timing.Truncated := TRUE;
   ELSE
       #Core.Timing.Rows[#Slot].Id := #Core.Command;
       #Core.Timing.Rows[#Slot].Label := #Core.CommandLabel;
       IF #Core.Timing.Rows[#Slot].Count < UDINT#4294967295 THEN
           #Core.Timing.Rows[#Slot].Count := #Core.Timing.Rows[#Slot].Count + 1;
       END_IF;
       #Core.Timing.Rows[#Slot].Last := #Core.Timing.LastCmdTime;
       IF #Core.Timing.Rows[#Slot].Count = 1 OR #Core.Timing.LastCmdTime < #Core.Timing.Rows[#Slot].Minimum THEN
           #Core.Timing.Rows[#Slot].Minimum := #Core.Timing.LastCmdTime;
       END_IF;
       IF #Core.Timing.LastCmdTime > #Core.Timing.Rows[#Slot].Maximum THEN
           #Core.Timing.Rows[#Slot].Maximum := #Core.Timing.LastCmdTime;
       END_IF;
       #AverageMs := DINT_TO_LINT(TIME_TO_DINT(#Core.Timing.Rows[#Slot].Avg));
       #AverageMs := #AverageMs + (UDINT_TO_LINT(#DurationMs) - #AverageMs) / UDINT_TO_LINT(#Core.Timing.Rows[#Slot].Count);
       #Core.Timing.Rows[#Slot].Avg := DINT_TO_TIME(LINT_TO_DINT(#AverageMs));
   END_IF;
   #Core.TimingOpen := FALSE;
END_FUNCTION

FUNCTION "FRK_ReleaseCommand" : Void   // FC19, SCL
{ S7_Optimized_Access := 'TRUE' }
VERSION : 0.1
// stored: AutoNumber true, IsIECCheckEnabled false, SetENOAutomatically false, UDAEnableTagReadback false
   VAR_IN_OUT
      Core : "FRK_Core";
      Execute : Bool;
   END_VAR
BEGIN

   #Execute := FALSE;
   #Core.ReleasePending := TRUE;
END_FUNCTION

FUNCTION "FRK_ReleaseReason" : Void   // FC43, SCL
{ S7_Optimized_Access := 'TRUE' }
VERSION : 0.1
// stored: AutoNumber true, IsIECCheckEnabled false, SetENOAutomatically false, UDAEnableTagReadback false
   VAR_INPUT
      Description : WString;
      Reason : DInt;
      Path : WString;
      Kind : DInt;
   END_VAR
   VAR_IN_OUT
      Report : "ST_ReleaseReport";
   END_VAR
BEGIN

   #Report.Released := FALSE;
   IF #Report.Count < 24 THEN
       #Report.Count := #Report.Count + 1;
       #Report.Reasons[#Report.Count].Description := #Description;
       #Report.Reasons[#Report.Count].ReasonCode := #Reason;
       #Report.Reasons[#Report.Count].SourcePath := #Path;
       #Report.Reasons[#Report.Count].Kind := #Kind;
       #Report.Reasons[#Report.Count].Bypassable := FALSE;
   END_IF;
END_FUNCTION

FUNCTION "FRK_Release_DeclarationUnit" : Void   // FC71, SCL
{ S7_Optimized_Access := 'TRUE' }
VERSION : 0.1
// stored: AutoNumber true, IsIECCheckEnabled false, SetENOAutomatically false, UDAEnableTagReadback false
   VAR_IN_OUT
      Unit : "FRK_Unit";
      Hal : "ST_DeclarationUnitHal";
   END_VAR
BEGIN

   "FRK_UnitSetPermit"(Unit := #Unit,
                       Ok := #Hal.Cell.Clamp.Permit,
                       Diag := #Hal.Cell.Clamp.Diag);
END_FUNCTION

FUNCTION "FRK_Release_InnerUnit" : Void   // FC65, SCL
{ S7_Optimized_Access := 'TRUE' }
VERSION : 0.1
// stored: AutoNumber true, IsIECCheckEnabled false, SetENOAutomatically false, UDAEnableTagReadback false
   VAR_IN_OUT
      Unit : "FRK_Unit";
      Hal : "ST_InnerUnitHal";
   END_VAR
BEGIN

   "FRK_UnitSetPermit"(Unit := #Unit,
                       Ok := #Hal.Cell.Clamp.Permit,
                       Diag := #Hal.Cell.Clamp.Diag);
END_FUNCTION

FUNCTION "FRK_Release_SatelliteUnit" : Void   // FC68, SCL
{ S7_Optimized_Access := 'TRUE' }
VERSION : 0.1
// stored: AutoNumber true, IsIECCheckEnabled false, SetENOAutomatically false, UDAEnableTagReadback false
   VAR_IN_OUT
      Unit : "FRK_Unit";
      Hal : "ST_SatelliteUnitHal";
   END_VAR
BEGIN

   "FRK_UnitSetPermit"(Unit := #Unit,
                       Ok := #Hal.Cell.Clamp.Permit,
                       Diag := #Hal.Cell.Clamp.Diag);
END_FUNCTION

FUNCTION "FRK_RouteAbort" : Void   // FC16, SCL
{ S7_Optimized_Access := 'TRUE' }
VERSION : 0.1
// stored: AutoNumber true, IsIECCheckEnabled false, SetENOAutomatically false, UDAEnableTagReadback false
   VAR_INPUT
      Abort : Bool;
   END_VAR
   VAR_IN_OUT
      Core : "FRK_Core";
   END_VAR
   VAR_TEMP
      ErrorAbort : Bool;
   END_VAR
BEGIN

   IF (#Abort OR #Core.ReleasePending) AND #Core.Exec = 1 THEN
       #Core.Exec := 4;
       #Core.Step := 0;
       #Core.Dispatch := FALSE;
       #Core.EvAbort := TRUE;
   END_IF;
   #ErrorAbort := (#Abort OR #Core.ReleasePending) AND #Core.Exec = 3;
   #Core.EvAbortInError := #ErrorAbort AND NOT #Core.AbortPrev;
   #Core.AbortPrev := #ErrorAbort;
END_FUNCTION

FUNCTION "FRK_Route_DeclarationCell" : Bool   // FC63, SCL
{ S7_Optimized_Access := 'TRUE' }
VERSION : 0.1
// stored: AutoNumber true, IsIECCheckEnabled false, SetENOAutomatically false, UDAEnableTagReadback false
   VAR_INPUT
      Request : "ST_HmiRequest";
   END_VAR
   VAR_IN_OUT
      Module : "FB_DeclarationCell";
      Hal : "ST_DeclarationCellHal";
      Report : "ST_ReleaseReport";
   END_VAR
   VAR_TEMP
      RouteMatched : Bool;
      Index : Int;
   END_VAR
BEGIN

   #FRK_Route_DeclarationCell := FALSE;
   IF NOT "FRK_PathOwned"(OwnerPath := #Module.Status.Name, TargetPath := #Request.TargetPath) THEN
       RETURN;
   END_IF;
   IF #Request.TargetPath = STRING_TO_WSTRING(#Module.Status.Name) THEN
       FOR #Index := 1 TO 16 DO
           #Module.ManConditions[#Index].Used := FALSE;
       END_FOR;
       "FRK_ManualApply"(Core := #Module.Core,
                         Status := #Module.Status,
                         Request := #Request,
                         Commands := #Module.Catalog,
                         Count := #Module.CatalogCount,
                         Conditions := #Module.ManConditions,
                         Report := #Report,
                         Execute := #Module.Execute,
                         Command := #Module.Command,
                         ManualOwned := #Module.ManualOwned);
       #FRK_Route_DeclarationCell := TRUE;
       RETURN;
   END_IF;
   #RouteMatched := "FRK_Route_DeclarationCylinder"(Module := #Module.Clamp, Hal := #Hal.Clamp, Request := #Request, Report := #Report);
   #FRK_Route_DeclarationCell := #FRK_Route_DeclarationCell OR #RouteMatched;
   #RouteMatched := "FRK_Route_DeclarationCylinder"(Module := #Module.Gate, Hal := #Hal.Gate, Request := #Request, Report := #Report);
   #FRK_Route_DeclarationCell := #FRK_Route_DeclarationCell OR #RouteMatched;
END_FUNCTION

FUNCTION "FRK_Route_DeclarationCylinder" : Bool   // FC61, SCL
{ S7_Optimized_Access := 'TRUE' }
VERSION : 0.1
// stored: AutoNumber true, IsIECCheckEnabled false, SetENOAutomatically false, UDAEnableTagReadback false
   VAR_INPUT
      Request : "ST_HmiRequest";
   END_VAR
   VAR_IN_OUT
      Module : "FB_DeclarationCylinder";
      Hal : "ST_DeclarationLeafHal";
      Report : "ST_ReleaseReport";
   END_VAR
   VAR_TEMP
      RouteMatched : Bool;
      Index : Int;
   END_VAR
BEGIN

   #FRK_Route_DeclarationCylinder := FALSE;
   IF NOT "FRK_PathOwned"(OwnerPath := #Module.Status.Name, TargetPath := #Request.TargetPath) THEN
       RETURN;
   END_IF;
   IF #Request.TargetPath = STRING_TO_WSTRING(#Module.Status.Name) THEN
       FOR #Index := 1 TO 16 DO
           #Module.ManConditions[#Index].Used := FALSE;
       END_FOR;
       // ---- AUTHORED: OnManRelease
       "FRK_ManualCondition"(Conditions := #Module.ManConditions,
                             Slot := 1,
                             Value := 2,
                             Ok := #Hal.Permit,
                             Diag := #Hal.Diag,
                             Bypassable := FALSE);
       "FRK_ManualCondition"(Conditions := #Module.ManConditions,
                             Slot := 2,
                             Value := 2,
                             Ok := #Hal.Sample = 0,
                             Diag := #Hal.LaterDiag,
                             Bypassable := FALSE);
       // ---- GENERATED: manual release end
       "FRK_ManualApply"(Core := #Module.Core,
                         Status := #Module.Status,
                         Request := #Request,
                         Commands := #Module.Catalog,
                         Count := #Module.CatalogCount,
                         Conditions := #Module.ManConditions,
                         Report := #Report,
                         Execute := #Module.Execute,
                         Command := #Module.Command,
                         ManualOwned := #Module.ManualOwned);
       #FRK_Route_DeclarationCylinder := TRUE;
       RETURN;
   END_IF;
END_FUNCTION

FUNCTION "FRK_Route_DeclarationUnit" : Bool   // FC72, SCL
{ S7_Optimized_Access := 'TRUE' }
VERSION : 0.1
// stored: AutoNumber true, IsIECCheckEnabled false, SetENOAutomatically false, UDAEnableTagReadback false
   VAR_INPUT
      Request : "ST_HmiRequest";
   END_VAR
   VAR_IN_OUT
      Module : "FB_DeclarationUnit";
      Hal : "ST_DeclarationUnitHal";
      Report : "ST_ReleaseReport";
   END_VAR
   VAR_TEMP
      RouteMatched : Bool;
      Index : Int;
   END_VAR
BEGIN

   #FRK_Route_DeclarationUnit := FALSE;
   IF NOT "FRK_PathOwned"(OwnerPath := #Module.Status.Name, TargetPath := #Request.TargetPath) THEN
       RETURN;
   END_IF;
   "FRK_Release_DeclarationUnit"(Unit := #Module.Unit,
                                 Hal := #Hal);
   "FRK_ManualCommon"(Core := #Module.Core,
                      Unit := #Module.Unit,
                      Status := #Module.Status,
                      Report := #Report);
   IF #Request.TargetPath = STRING_TO_WSTRING(#Module.Status.Name) THEN
       "FRK_ReleaseReason"(Report := #Report,
                           Description := WSTRING#'std.error.unsupportedHmiRequest',
                           Reason := 2008,
                           Path := STRING_TO_WSTRING(#Module.Status.Name),
                           Kind := 4);
       #FRK_Route_DeclarationUnit := TRUE;
       RETURN;
   END_IF;
   #RouteMatched := "FRK_Route_DeclarationCell"(Module := #Module.Cell, Hal := #Hal.Cell, Request := #Request, Report := #Report);
   #FRK_Route_DeclarationUnit := #FRK_Route_DeclarationUnit OR #RouteMatched;
   #RouteMatched := "FRK_Route_SatelliteUnit"(Module := #Module.Satellite, Hal := #Hal.Satellite, Request := #Request, Report := #Report);
   #FRK_Route_DeclarationUnit := #FRK_Route_DeclarationUnit OR #RouteMatched;
END_FUNCTION

FUNCTION "FRK_Route_InnerUnit" : Bool   // FC66, SCL
{ S7_Optimized_Access := 'TRUE' }
VERSION : 0.1
// stored: AutoNumber true, IsIECCheckEnabled false, SetENOAutomatically false, UDAEnableTagReadback false
   VAR_INPUT
      Request : "ST_HmiRequest";
   END_VAR
   VAR_IN_OUT
      Module : "FB_InnerUnit";
      Hal : "ST_InnerUnitHal";
      Report : "ST_ReleaseReport";
   END_VAR
   VAR_TEMP
      RouteMatched : Bool;
      Index : Int;
   END_VAR
BEGIN

   #FRK_Route_InnerUnit := FALSE;
   IF NOT "FRK_PathOwned"(OwnerPath := #Module.Status.Name, TargetPath := #Request.TargetPath) THEN
       RETURN;
   END_IF;
   "FRK_Release_InnerUnit"(Unit := #Module.Unit,
                           Hal := #Hal);
   "FRK_ManualCommon"(Core := #Module.Core,
                      Unit := #Module.Unit,
                      Status := #Module.Status,
                      Report := #Report);
   IF #Request.TargetPath = STRING_TO_WSTRING(#Module.Status.Name) THEN
       "FRK_ReleaseReason"(Report := #Report,
                           Description := WSTRING#'std.error.unsupportedHmiRequest',
                           Reason := 2008,
                           Path := STRING_TO_WSTRING(#Module.Status.Name),
                           Kind := 4);
       #FRK_Route_InnerUnit := TRUE;
       RETURN;
   END_IF;
   #RouteMatched := "FRK_Route_DeclarationCell"(Module := #Module.Cell, Hal := #Hal.Cell, Request := #Request, Report := #Report);
   #FRK_Route_InnerUnit := #FRK_Route_InnerUnit OR #RouteMatched;
END_FUNCTION

FUNCTION "FRK_Route_SatelliteUnit" : Bool   // FC69, SCL
{ S7_Optimized_Access := 'TRUE' }
VERSION : 0.1
// stored: AutoNumber true, IsIECCheckEnabled false, SetENOAutomatically false, UDAEnableTagReadback false
   VAR_INPUT
      Request : "ST_HmiRequest";
   END_VAR
   VAR_IN_OUT
      Module : "FB_SatelliteUnit";
      Hal : "ST_SatelliteUnitHal";
      Report : "ST_ReleaseReport";
   END_VAR
   VAR_TEMP
      RouteMatched : Bool;
      Index : Int;
   END_VAR
BEGIN

   #FRK_Route_SatelliteUnit := FALSE;
   IF NOT "FRK_PathOwned"(OwnerPath := #Module.Status.Name, TargetPath := #Request.TargetPath) THEN
       RETURN;
   END_IF;
   "FRK_Release_SatelliteUnit"(Unit := #Module.Unit,
                               Hal := #Hal);
   "FRK_ManualCommon"(Core := #Module.Core,
                      Unit := #Module.Unit,
                      Status := #Module.Status,
                      Report := #Report);
   IF #Request.TargetPath = STRING_TO_WSTRING(#Module.Status.Name) THEN
       "FRK_ReleaseReason"(Report := #Report,
                           Description := WSTRING#'std.error.unsupportedHmiRequest',
                           Reason := 2008,
                           Path := STRING_TO_WSTRING(#Module.Status.Name),
                           Kind := 4);
       #FRK_Route_SatelliteUnit := TRUE;
       RETURN;
   END_IF;
   #RouteMatched := "FRK_Route_DeclarationCell"(Module := #Module.Cell, Hal := #Hal.Cell, Request := #Request, Report := #Report);
   #FRK_Route_SatelliteUnit := #FRK_Route_SatelliteUnit OR #RouteMatched;
   #RouteMatched := "FRK_Route_InnerUnit"(Module := #Module.Inner, Hal := #Hal.Inner, Request := #Request, Report := #Report);
   #FRK_Route_SatelliteUnit := #FRK_Route_SatelliteUnit OR #RouteMatched;
END_FUNCTION

FUNCTION "FRK_SetIdentity" : Void   // FC1, SCL
{ S7_Optimized_Access := 'TRUE' }
VERSION : 0.1
// Generated registry services v0.1; compact rows contain no operator strings.
// stored: AutoNumber true, IsIECCheckEnabled false, SetENOAutomatically false, UDAEnableTagReadback false
   VAR_INPUT
      InstancePath : WString;
      ModuleType : DInt;
      TypeId : DInt;
      Capabilities : DWord;
      ParentIndex : DInt;
      TypeKey : String;
   END_VAR
   VAR_IN_OUT
      Core : "FRK_Core";
      Status : "ST_ModuleStatus";
   END_VAR
   VAR_TEMP
      Identity : String[254];
      QuotePos : Int;
      RowIndex : DInt;
   END_VAR
BEGIN

